(* IEC 61131-3 sources: volt/packages/volt-lsp-iec/test-corpus/bakon-nano/Device/Plc Logic/Application/Library Manager/L_MC1P_MotionControlBasic (part 2) *)

(* ---- L_MC1P_IAXISCOMMMAND.itf ---- *)
INTERFACE L_MC1P_IAXISCOMMMAND
END_INTERFACE

METHOD ABORTING
END_METHOD

METHOD CALCSTATUS
VAR_IN_OUT
	AXIS : _AXIS_REF_REAL;
END_VAR
END_METHOD

METHOD EXECUTE
END_METHOD

METHOD MAIN
END_METHOD

METHOD RESETCOMMANDERRORSTATE : BOOL
VAR_IN_OUT
	AXIS : _AXIS_REF_REAL;
END_VAR
END_METHOD

METHOD RESETSTATUSPARAMETER
END_METHOD

METHOD SETINCTANCEINFO
VAR_INPUT
	PSINSTANCENAME : POINTER TO STRING;
	ERRORITFID : DWORD;
END_VAR
END_METHOD

METHOD UPDATEAXISPOINTER
VAR_INPUT
	PAXIS : POINTER TO AXIS_REF;
END_VAR
END_METHOD

METHOD UPDATECOMMANDINTERFACE
VAR_IN_OUT
	CMD : USINT;
END_VAR
END_METHOD

(* ---- L_MC1P_IAXISCOMMMAND_AUTOTUNING.itf ---- *)
INTERFACE L_MC1P_IAXISCOMMMAND_AUTOTUNING
END_INTERFACE

METHOD CALCPROFILEPARAMS
VAR_IN_OUT
	AXIS : AXIS_REF;
END_VAR
END_METHOD

METHOD UPDATEPARAINTERFACE
VAR_IN_OUT
	SCPAR : L_MC1P_AutotuningPara;
END_VAR
END_METHOD

(* ---- L_MC1P_IAXISEXTENSION.itf ---- *)
INTERFACE L_MC1P_IAXISEXTENSION
END_INTERFACE

METHOD SETBASICINITIALISATION
VAR_INPUT
	ITFGENERICCONFIG : L_MC1P_IGenericAxisConfiguration;
END_VAR
VAR_IN_OUT
	AXIS : _AXIS_REF_REAL;
END_VAR
END_METHOD

(* ---- L_MC1P_IAXISSIMCALLSINGLESTEPS.itf ---- *)
INTERFACE L_MC1P_IAXISSIMCALLSINGLESTEPS
END_INTERFACE

METHOD SIMFINISH : BOOL
VAR_INPUT
	AXISID : INT;
	ITFMECHANICSIMULATION : L_MC1P_IMechanicSimulation;
END_VAR
VAR_IN_OUT
	AXIS : _AXIS_REF_REAL;
END_VAR
END_METHOD

METHOD SIMINSIDELOOP : BOOL
VAR_INPUT
	AXISID : INT;
	ISYSTEMSIMCOUNTER : INT;
	ITFMECHANICSIMULATION : L_MC1P_IMechanicSimulation;
END_VAR
END_METHOD

METHOD SIMPREPARE : BOOL
VAR_INPUT
	AXISID : INT;
	ITFMECHANICSIMULATION : L_MC1P_IMechanicSimulation;
END_VAR
VAR_IN_OUT
	AXIS : _AXIS_REF_REAL;
END_VAR
END_METHOD

(* ---- L_MC1P_IAXISSIMULATIONINTERFACE.itf ---- *)
INTERFACE L_MC1P_IAXISSIMULATIONINTERFACE
END_INTERFACE

METHOD ACTIVATESIMULATION
VAR_IN_OUT
	AXIS : _AXIS_REF_REAL;
END_VAR
END_METHOD

METHOD CALCULATEINPUTDATA
VAR_INPUT
	ITFKINSIM : L_MC1P_IKinematicSimulation;
END_VAR
VAR_IN_OUT
	AXIS : _AXIS_REF_REAL;
END_VAR
END_METHOD

METHOD CALCULATEOUTPUTDATA
VAR_INPUT
	ITFKINSIM : L_MC1P_IKinematicSimulation;
END_VAR
VAR_IN_OUT
	AXIS : _AXIS_REF_REAL;
END_VAR
END_METHOD

METHOD DISABLESIMULATION
VAR_IN_OUT
	AXIS : _AXIS_REF_REAL;
END_VAR
END_METHOD

(* ---- L_MC1P_ICOMMMUNICATIONSIMULATION.itf ---- *)
INTERFACE L_MC1P_ICOMMMUNICATIONSIMULATION
END_INTERFACE

METHOD GETCOMMSTATE : L_DCO_CommState
VAR_INPUT
	PAXISCOMM : POINTER TO _AXIS_REF_COM;
END_VAR
END_METHOD

METHOD PARREAD
VAR_INPUT
	WIDX : DWORD;
END_VAR
END_METHOD

METHOD PARREAD_GETOUTPUT
VAR_INPUT
	WIDX : DWORD;
END_VAR
VAR_OUTPUT
	SZDATAREAD : CAA_SIZE;
	XDONE : BOOL;
	XERROR : BOOL;
	WERROR : WORD;
END_VAR
END_METHOD

METHOD PARREAD_SETINPUT
VAR_INPUT
	WIDX : DWORD;
	XEXECUTE : BOOL;
	WINDEX : WORD;
	BYSUBINDEX : BYTE;
	PBUFFER : POINTER TO BYTE;
	SZSIZE : UDINT;
	UDITIMEOUT : UDINT;
	XSLOTB : BOOL;
END_VAR
END_METHOD

METHOD PARWRITE
VAR_INPUT
	WIDX : DWORD;
END_VAR
END_METHOD

METHOD PARWRITE_GETOUTPUT
VAR_INPUT
	WIDX : DWORD;
END_VAR
VAR_OUTPUT
	XDONE : BOOL;
	XERROR : BOOL;
	WERROR : WORD;
END_VAR
END_METHOD

METHOD PARWRITE_SETINPUT
VAR_INPUT
	WIDX : DWORD;
	XEXECUTE : BOOL;
	WINDEX : WORD;
	BYSUBINDEX : BYTE;
	PBUFFER : POINTER TO BYTE;
	SZSIZE : UDINT;
	UDITIMEOUT : UDINT;
	XSLOTB : BOOL;
END_VAR
END_METHOD

METHOD RESTARTMASTER
VAR_INPUT
	XEXECUTE : BOOL;
	PAXIS : POINTER TO _AXIS_REF_COM;
END_VAR
VAR_OUTPUT
	XDONE : BOOL;
	XERROR : BOOL;
	XBUSY : BOOL;
	DWERROR : DWORD;
END_VAR
END_METHOD

(* ---- L_MC1P_ICOMMUNICATION.itf ---- *)
INTERFACE L_MC1P_ICOMMUNICATION
END_INTERFACE

METHOD FORWARDERROR
VAR_INPUT
	XENABLE : BOOL;
	XWARNING : BOOL;
	XERROR : BOOL;
	WERRORID : WORD;
	WTEXTREFID : WORD;
	XRESETERROR : BOOL := FALSE;
	AXISMODULEHANDLER : L_IMHP_IModuleHandler;
END_VAR
END_METHOD

METHOD GETCOMMPARAMETER
VAR_INPUT
	PCONNECTOR : POINTER TO IoConfigConnector;
END_VAR
VAR_OUTPUT
	PSLAVECONNECTOR : POINTER TO IoStandard.IoConfigConnector;
	UINETID : UINT;
	UIDEVICEID : UINT;
	XSENDFRAMEATTASKSTART : BOOL;
	UDIPRODUCTCODE : DWORD;
	PMASTERCONNECTOR : POINTER TO IoStandard.IoConfigConnector;
END_VAR
END_METHOD

METHOD GETCOMMSTATE : L_DCO_CommState
VAR_INPUT
	PAXISCOMM : POINTER TO _AXIS_REF_COM;
END_VAR
END_METHOD

METHOD GETPDINEQPDOUT : BOOL
END_METHOD

METHOD PARREAD
VAR_INPUT
	WIDX : DWORD;
END_VAR
END_METHOD

METHOD PARREAD_GETOUTPUT
VAR_INPUT
	WIDX : DWORD;
END_VAR
VAR_OUTPUT
	SZDATAREAD : CAA_SIZE;
	XDONE : BOOL;
	XERROR : BOOL;
	WERROR : WORD;
END_VAR
END_METHOD

METHOD PARREAD_SETINPUT
VAR_INPUT
	WIDX : DWORD;
	XEXECUTE : BOOL;
	WINDEX : WORD;
	BYSUBINDEX : BYTE;
	PBUFFER : POINTER TO BYTE;
	SZSIZE : UDINT;
	UDITIMEOUT : UDINT;
END_VAR
END_METHOD

METHOD PARWRITE
VAR_INPUT
	WIDX : DWORD;
END_VAR
END_METHOD

METHOD PARWRITE_GETOUTPUT
VAR_INPUT
	WIDX : DWORD;
END_VAR
VAR_OUTPUT
	XDONE : BOOL;
	XERROR : BOOL;
	WERROR : WORD;
END_VAR
END_METHOD

METHOD PARWRITE_SETINPUT
VAR_INPUT
	WIDX : DWORD;
	XEXECUTE : BOOL;
	WINDEX : WORD;
	BYSUBINDEX : BYTE;
	PBUFFER : POINTER TO BYTE;
	SZSIZE : UDINT;
	UDITIMEOUT : UDINT;
END_VAR
END_METHOD

METHOD RESET
END_METHOD

METHOD RESTARTMASTER
VAR_INPUT
	XEXECUTE : BOOL;
	PAXIS : POINTER TO _AXIS_REF_COM;
END_VAR
VAR_OUTPUT
	XDONE : BOOL;
	XERROR : BOOL;
	XBUSY : BOOL;
	DWERROR : DWORD;
END_VAR
END_METHOD

METHOD SETBASICINITIALISATION
VAR_IN_OUT
	AXIS : _AXIS_REF_REAL;
END_VAR
END_METHOD

METHOD SETCOMPONENTINFO
VAR_INPUT
	DATASELECTION : WORD;
	SDATA : STRING;
END_VAR
END_METHOD

(* ---- L_MC1P_ICOMPENSATIONINTERFACE.itf ---- *)
INTERFACE L_MC1P_ICOMPENSATIONINTERFACE
END_INTERFACE

METHOD GETOFFSETVALUES
VAR_OUTPUT
	LROFFSETPOS : LREAL;
	LROFFSETVEL : LREAL;
	LROFFSETACC : LREAL;
END_VAR
END_METHOD

(* ---- L_MC1P_ICONFIGUREDRIVE.itf ---- *)
INTERFACE L_MC1P_ICONFIGUREDRIVE
END_INTERFACE

METHOD DOFUNCTION : BOOL
VAR_INPUT
	XEXECUTE : BOOL;
	WOFFSET : WORD;
END_VAR
VAR_OUTPUT
	XDONE : BOOL;
	XERROR : BOOL;
	XBUSY : BOOL;
	EERRORID : WORD;
END_VAR
VAR_IN_OUT
	AXIS : _AXIS_REF_REAL;
END_VAR
END_METHOD

METHOD GETADDITIONALCONFIGINFO : POINTER TO L_MC1P_AdditionalConfigInfo
END_METHOD

METHOD GETINSTANCE : POINTER TO BYTE
END_METHOD

METHOD RESET : BOOL
END_METHOD

(* ---- L_MC1P_ICONTROLLERADAPTION.itf ---- *)
INTERFACE L_MC1P_ICONTROLLERADAPTION
END_INTERFACE

METHOD CALCADAPTIONCURVE : LREAL
VAR_INPUT
	LRSETVEL : LREAL;
END_VAR
VAR_IN_OUT
	AXIS : _AXIS_REF_REAL;
END_VAR
END_METHOD

(* ---- L_MC1P_ICONTROLLERINTERFACE.itf ---- *)
INTERFACE L_MC1P_ICONTROLLERINTERFACE
END_INTERFACE

METHOD CALCCONTROLLER
VAR_INPUT
	LRSETPOSITION : LREAL;
	LRSETVELOCITY : LREAL;
	LRSETACCELERATION : LREAL;
	LRSETTORQUE : LREAL;
	LRSETJERK : LREAL;
	LRACTPOSITIONIN : LREAL;
	LRACTVELOCITYIN : LREAL;
	LRACTACCELERATIONIN : LREAL;
	LRACTTORQUEIN : LREAL;
END_VAR
VAR_OUTPUT
	LRSETPOSITIONOUT : LREAL;
	LRSETVELOCITYOUT : LREAL;
	LRSETACCELERATIONOUT : LREAL;
	LRSETTORQUEOUT : LREAL;
END_VAR
VAR_IN_OUT
	AXIS : _AXIS_REF_REAL;
END_VAR
END_METHOD

(* ---- L_MC1P_IDRIVESCALING.itf ---- *)
INTERFACE L_MC1P_IDRIVESCALING
END_INTERFACE

METHOD CALCACCFACTOR : BOOL
VAR_OUTPUT
	LRSCALEUNITTOACC : LREAL;
	LRSCALEACCTOUNIT : LREAL;
END_VAR
VAR_IN_OUT
	AXIS : _AXIS_REF_REAL;
END_VAR
END_METHOD

METHOD CALCSPEEDFACTOR : BOOL
VAR_OUTPUT
	LRSCALEUNITTOSPEED : LREAL;
	LRSCALESPEEDTOUNIT : LREAL;
END_VAR
VAR_IN_OUT
	AXIS : _AXIS_REF_REAL;
END_VAR
END_METHOD

METHOD CALCTORQUEFACTOR : BOOL
VAR_OUTPUT
	LRSCALETORQUETONORM : LREAL;
	LRSCALETORQUETONORM2 : LREAL;
	LRSCALENORMTOTORQUE : LREAL;
END_VAR
VAR_IN_OUT
	AXIS : _AXIS_REF_REAL;
END_VAR
END_METHOD

METHOD CHECKVALIDPOSRESOLUTION : BOOL
VAR_INPUT
	DWPOSRESOLUTION : DWORD;
END_VAR
END_METHOD

METHOD GETDEFAULTTORQUE : LREAL
VAR_INPUT
	LRREFTORQUE : LREAL;
END_VAR
END_METHOD

METHOD POSDIFFTOSPEEDINC : DINT
VAR_INPUT
	DIPOSDIFF : DINT := 0;
	DWFACTOR : DWORD := 1000;
END_VAR
VAR_IN_OUT
	AXIS : _AXIS_REF_REAL;
END_VAR
END_METHOD

METHOD SPEEDTOPOSDIFFINC : DINT
VAR_INPUT
	DISPEED : DINT := 0;
	DWFACTOR : DWORD := 1000;
END_VAR
VAR_IN_OUT
	AXIS : _AXIS_REF_REAL;
	DIRES : DINT;
END_VAR
END_METHOD

(* ---- L_MC1P_IDRIVESPECIFICIMPLBASE.itf ---- *)
INTERFACE L_MC1P_IDRIVESPECIFICIMPLBASE
END_INTERFACE

METHOD CALCAFTERREADINPUTS
VAR_IN_OUT
	AXIS : _AXIS_REF_REAL;
END_VAR
END_METHOD

METHOD CALCBEFOREREADINPUTS
VAR_IN_OUT
	AXIS : _AXIS_REF_REAL;
END_VAR
END_METHOD

METHOD CALCBEFOREWRITEOUTPUTS
VAR_IN_OUT
	AXIS : _AXIS_REF_REAL;
END_VAR
END_METHOD

METHOD CHECKAVAILABLECONTROLMODE : BOOL
VAR_IN_OUT
	AXIS : _AXIS_REF_REAL;
	POSCTRLDRIVEAVAILABLE : L_IE1P_Error;
	POSCTRLPLCAVAILABLE : L_IE1P_Error;
	SPEEDCTRLDRIVEAVAILABLE : L_IE1P_Error;
	TORQUECTRLDRIVE : L_IE1P_Error;
END_VAR
END_METHOD

METHOD CHECKRESETHOMEPOS
VAR_INPUT
	WFDBSTATUSWORD : WORD;
END_VAR
VAR_IN_OUT
	AXIS : _AXIS_REF_REAL;
END_VAR
END_METHOD

METHOD CHECKSAFETYOPTIONAVAILABLE : BOOL
VAR_INPUT
	DWPRODUCTCODE : DWORD;
END_VAR
END_METHOD

METHOD COLLECTDRIVESTATE : BOOL
VAR_IN_OUT
	AXIS : _AXIS_REF_REAL;
	SCSTATEINFO : L_MC1P_DriveStateCollection;
END_VAR
END_METHOD

METHOD CONTROLDRIVE : BOOL
VAR_INPUT
	XENABLE : BOOL;
END_VAR
VAR_IN_OUT
	AXIS : _AXIS_REF_REAL;
END_VAR
END_METHOD

METHOD DRIVECONFIGDATA
VAR_INPUT
	PCONFIGINFO : POINTER TO L_MC1P_AdditionalConfigInfo;
END_VAR
VAR_IN_OUT
	AXIS : _AXIS_REF_REAL;
END_VAR
END_METHOD

METHOD DRIVEFAULTSTATUS : BOOL
VAR_IN_OUT
	AXIS : _AXIS_REF_REAL;
	SCSTATEINFO : L_MC1P_DriveStateCollection;
END_VAR
END_METHOD

METHOD GETBRAKE : POINTER TO L_MC1P_BrakeControlBase
VAR_IN_OUT
	AXIS : _AXIS_REF_REAL;
END_VAR
END_METHOD

METHOD GETBRAKESERVICE : POINTER TO L_MC1P_BrakeService
VAR_IN_OUT
	AXIS : _AXIS_REF_REAL;
END_VAR
END_METHOD

METHOD GETCAUSEOFCINH : WORD
VAR_IN_OUT
	AXIS : _AXIS_REF_REAL;
END_VAR
END_METHOD

METHOD GETFDBSTATUSWORD : WORD
VAR_IN_OUT
	AXIS : _AXIS_REF_REAL;
END_VAR
END_METHOD

METHOD GETIECADRESS : BOOL
VAR_IN_OUT
	AXIS : _AXIS_REF_REAL;
	M_PPDOINFOCONNECTOR : POINTER TO IoConfigConnector;
	ATRANSELEMENT : ARRAY [1.._AXIS_REF_REAL.c_wMaxTransElem] OF L_MC1P_MappedElement;
	WTRANSELEMENTS : WORD;
	LWTRANSDATA : LWORD;
	LWRECDATA : LWORD;
	WRECEIVEELEMENTS : WORD;
	ARECEIVEELEMENT : ARRAY [1.._AXIS_REF_REAL.c_wMaxRecElem] OF L_MC1P_MappedElement;
END_VAR
END_METHOD

METHOD GETOPTIONALACTVEL : BOOL
VAR_IN_OUT
	LRVEL : LREAL;
END_VAR
END_METHOD

METHOD GETRECEIVEDATAIMPL : DWORD
VAR_INPUT
	LWMASK : LWORD;
END_VAR
VAR_IN_OUT
	AXIS : _AXIS_REF_REAL;
END_VAR
END_METHOD

METHOD GETSTATUSWORDS
VAR_OUTPUT
	STATUSWORD1 : WORD;
	STATUSWORD2 : WORD;
	STATUSWORD3 : WORD;
	STATUSWORD4 : WORD;
END_VAR
VAR_IN_OUT
	AXIS : _AXIS_REF_REAL;
END_VAR
END_METHOD

METHOD GETTRANSMITDATAIMPL : DWORD
VAR_INPUT
	LWMASK : LWORD;
END_VAR
VAR_IN_OUT
	AXIS : _AXIS_REF_REAL;
END_VAR
END_METHOD

METHOD GETTRANSMITDATALREALIMPL : LREAL
VAR_INPUT
	LWMASK : LWORD;
END_VAR
VAR_IN_OUT
	AXIS : _AXIS_REF_REAL;
END_VAR
END_METHOD

METHOD HOMECONFIG : BOOL
VAR_INPUT
	LRPOSITION : LREAL;
END_VAR
VAR_OUTPUT
	WINDEX : WORD;
	BYSUBINDEX : BYTE;
	BYNROFBYTE : BYTE;
	DWDATA : DWORD;
	XWRITEPARAM : BOOL;
	XDONE : BOOL;
	XERROR : BOOL;
END_VAR
VAR_IN_OUT
	AXIS : _AXIS_REF_REAL;
	SCHOMEDATA : L_MC1P_HomeParameter;
	WSTEP : WORD;
END_VAR
END_METHOD

METHOD HOMEPOSPERMANENTSETACTIVE : BOOL
VAR_IN_OUT
	AXIS : _AXIS_REF_REAL;
END_VAR
END_METHOD

METHOD RECEIVEPARAMETER
VAR_INPUT
	WPARAMETER : WORD;
	PADRESS : POINTER TO BYTE;
	WSIZE : WORD;
END_VAR
VAR_IN_OUT
	AXIS : _AXIS_REF_REAL;
END_VAR
END_METHOD

METHOD RECEIVEPARAMETERCALC
VAR_IN_OUT
	AXIS : _AXIS_REF_REAL;
	DATA : ARRAY [1..L_MC1P_Constants.gc_Rec_MaxDataIndex] OF POINTER TO L_MC1P_MappedElement;
END_VAR
END_METHOD

METHOD RESETDRIVECONTROL
VAR_INPUT
	XRESETDRIVEERROR : BOOL;
END_VAR
END_METHOD

METHOD RESTOREADDITIONALRETAINDATA
VAR_INPUT
	PDATA : POINTER TO L_MC1P_uRetainData;
END_VAR
END_METHOD

METHOD SETAXISPROPERTIES
VAR_IN_OUT
	AXIS : _AXIS_REF_REAL;
	AXISPROPERTIES : L_MC1P_AxisProperties;
END_VAR
END_METHOD

METHOD SETAXISSTATUSWORD
VAR_IN_OUT
	AXIS : _AXIS_REF_REAL;
	DWAXISSTATUS : DWORD;
END_VAR
END_METHOD

METHOD SETBASICINITIALISATION
VAR_IN_OUT
	AXIS : _AXIS_REF_REAL;
END_VAR
END_METHOD

METHOD SETCONTROLWORDS
VAR_INPUT
	CONTROLWORD1 : WORD;
	CONTROLWORD2 : WORD;
	CONTROLWORD3 : WORD;
	CONTROLWORD4 : WORD;
END_VAR
VAR_IN_OUT
	AXIS : _AXIS_REF_REAL;
END_VAR
END_METHOD

METHOD SETDCBRAKE
VAR_INPUT
	XSETDCBRAKE : BOOL;
END_VAR
VAR_OUTPUT
	XDCBRAKEACTIVE : BOOL;
END_VAR
VAR_IN_OUT
	AXIS : _AXIS_REF_REAL;
END_VAR
END_METHOD

METHOD SETDRIVECONFIGINIT
VAR_IN_OUT
	AXIS : _AXIS_REF_REAL;
END_VAR
END_METHOD

METHOD SETSPEEDCTRLLIMITATION : BOOL
VAR_INPUT
	XLIMIT : BOOL;
END_VAR
VAR_IN_OUT
	AXIS : _AXIS_REF_REAL;
END_VAR
END_METHOD

METHOD SETSPEEDCTRLLOADVALUE
VAR_INPUT
	XLOAD : BOOL;
	LRVALUE : LREAL;
END_VAR
VAR_IN_OUT
	AXIS : _AXIS_REF_REAL;
END_VAR
END_METHOD

METHOD STOREADDITIONALRETAINDATA
VAR_INPUT
	PDATA : POINTER TO L_MC1P_uRetainData;
END_VAR
END_METHOD

METHOD TRANSMITPARAMETER
VAR_INPUT
	WPARAMETER : WORD;
	PADRESS : POINTER TO BYTE;
	WSIZE : WORD;
END_VAR
VAR_IN_OUT
	AXIS : _AXIS_REF_REAL;
END_VAR
END_METHOD

METHOD TRANSMITPARAMETERCALC
VAR_IN_OUT
	AXIS : _AXIS_REF_REAL;
	DATA : ARRAY [1..L_MC1P_Constants.gc_Trans_MaxDataIndex] OF POINTER TO L_MC1P_MappedElement;
END_VAR
END_METHOD

METHOD UPDATEMAPPING
VAR_INPUT
	PTASKMAPLIST : POINTER TO IoStandard.IoConfigTaskMap;
	NCOUNT : DINT;
	PPDOINFOCONNECTOR : POINTER TO IoConfigConnector;
END_VAR
VAR_IN_OUT
	AXIS : _AXIS_REF_REAL;
END_VAR
END_METHOD

(* ---- L_MC1P_IDRIVEUTILS.itf ---- *)
INTERFACE L_MC1P_IDRIVEUTILS
END_INTERFACE

METHOD ACTIVATEAPPCREDITS
VAR_INPUT
	XACTIVATE : BOOL;
END_VAR
END_METHOD

METHOD GETMULTIAXISINFO
VAR_IN_OUT
	MULTIAXISINFO : L_MC1P_MultiAxisInfo;
END_VAR
END_METHOD

METHOD GETRETAINMEMINFO : L_MC1P_RetainDataType
VAR_OUTPUT
	MEMINFO : L_MC1P_uAxisRetainInfo;
END_VAR
END_METHOD

METHOD RESETCONNECTION : L_IE1P_Error
VAR_INPUT
	ITFCALLEDFUNCITON : L_IF1P_IFunctionConnection;
	EDISCONNECTMODE : L_IF1P_DisconnectMode;
	XDISCONNECTEXISTINGCONNECTION : BOOL;
END_VAR
END_METHOD

METHOD SETCONNECTION
VAR_INPUT
	AXISCONNECTION : L_IF1P_IFunctionConnection;
END_VAR
END_METHOD

(* ---- L_MC1P_IENCODERINTERFACE.itf ---- *)
INTERFACE L_MC1P_IENCODERINTERFACE
END_INTERFACE

METHOD ENCNEWHOMEPOSLOADED : BOOL
VAR_INPUT
	DWCALLYCLE : DWORD;
	DWDELAY : DWORD;
END_VAR
END_METHOD

METHOD ENCRESETACTPOS
END_METHOD

METHOD ENCRESETHOMEPOS
VAR_INPUT
	ERESETINFO : L_IE1P_Error;
END_VAR
END_METHOD

METHOD ENCSETHOMEPOSITION
VAR_INPUT
	POSITION : LREAL;
	RELATIVE : BOOL;
	POSDIFF : LREAL;
	EHOMEPOSINFO : L_IE1P_Error;
END_VAR
END_METHOD

METHOD ENCSIGNALVALID : BOOL
VAR_OUTPUT
	XSIGNALVALIDOLD : BOOL;
	EENCERRORID : L_IE1P_Error;
END_VAR
END_METHOD

METHOD GETACTPOSINCR : DINT
END_METHOD

METHOD GETACTPOSINCR1616 : DINT
END_METHOD

METHOD GETACTVALUES
VAR_OUTPUT
	LRACTPOS : LREAL;
	LRACTVEL : LREAL;
	LRACTACC : LREAL;
	LRACTPOSUNFILTERED : LREAL;
	LRACTPOSROUNDS : LREAL;
END_VAR
END_METHOD

METHOD GETAXISINSTANCE : POINTER TO _AXIS_REF_REAL
END_METHOD

METHOD GETCONFIGCHANGED : BOOL
END_METHOD

METHOD GETHOMEPOSAVAILABLE : BOOL
END_METHOD

METHOD SETHOMEPOSAVAILABLE
VAR_INPUT
	XHOMEPOSAVAILABLE : BOOL;
END_VAR
END_METHOD

(* ---- L_MC1P_IENCODERPOSFILTER.itf ---- *)
INTERFACE L_MC1P_IENCODERPOSFILTER
END_INTERFACE

METHOD CALCULATE
VAR_INPUT
	LRCYCPOSIN : LREAL;
	LRCYCVELIN : LREAL;
END_VAR
VAR_OUTPUT
	LRCYCPOSOUT : LREAL;
	LRCYCVELOUT : LREAL;
	WFILTERSTATE : WORD;
END_VAR
END_METHOD

METHOD INIT
END_METHOD

METHOD RESET
END_METHOD

(* ---- L_MC1P_IERRORHANDLINGAXISSYSTEMS.itf ---- *)
INTERFACE L_MC1P_IERRORHANDLINGAXISSYSTEMS
END_INTERFACE

METHOD CLEARERRORINAXISSYSTEM
VAR_INPUT
	INSTANCEID : DWORD := 0;
END_VAR
END_METHOD

METHOD GETERRORITFID : DWORD
END_METHOD

METHOD NOTIFYERRORINAXISSYSTEM : BOOL
VAR_INPUT
	WERRORID : L_IE1P_Error := 0;
	INSTANCEID : DWORD := 0;
	PSINSTANCENAME : POINTER TO BYTE := 0;
	EERRORREACTION : L_IE1P_SeverityLevel := 0;
END_VAR
END_METHOD

(* ---- L_MC1P_IEXTENDEDMAPPINGACCESS.itf ---- *)
INTERFACE L_MC1P_IEXTENDEDMAPPINGACCESS
END_INTERFACE

METHOD GETIECADRESS
VAR_INPUT
	AXISCONNECTOR : POINTER TO IoConfigConnector;
END_VAR
END_METHOD

METHOD GETMAPPEDDATA : POINTER TO BYTE
VAR_INPUT
	UIINDEX : WORD;
	USISUBINDEX : USINT;
	USISIZE : USINT;
	XWRITEACCESS : BOOL;
	PADDDATA : POINTER TO BYTE;
	PXWAITFORINITACCESS : POINTER TO BOOL;
END_VAR
VAR_OUTPUT
	EERRORID : L_IE1P_Error;
	XERROR : BOOL;
	USISIZEACT : USINT;
END_VAR
END_METHOD

METHOD GETMAPPEDDATASUPPORT : BOOL
END_METHOD

METHOD RESETOUTPUTMAPPINGOBJECTS : BOOL
END_METHOD

(* ---- L_MC1P_IGENERICAXISCONFIGURATION.itf ---- *)
INTERFACE L_MC1P_IGENERICAXISCONFIGURATION
END_INTERFACE

METHOD CALCAFTERREADINPUTS
VAR_IN_OUT
	AXIS : _AXIS_REF_REAL;
	DRIVESPECIFIC : L_MC1P_DriveSpecific_Generic;
END_VAR
END_METHOD

METHOD CALCBEFOREREADINPUTS
VAR_IN_OUT
	AXIS : _AXIS_REF_REAL;
	DRIVESPECIFIC : L_MC1P_DriveSpecific_Generic;
END_VAR
END_METHOD

METHOD CALCBEFOREWRITEOUTPUTS
VAR_IN_OUT
	AXIS : _AXIS_REF_REAL;
	DRIVESPECIFIC : L_MC1P_DriveSpecific_Generic;
END_VAR
END_METHOD

METHOD DRIVECONFIG
VAR_INPUT
	WOFFSET : WORD;
END_VAR
VAR_OUTPUT
	XCONFIGBUSY : BOOL;
	XWAITFORPARAMETERWRITEDONE : BOOL;
	XWAITFORPARAMETERREADDONE : BOOL;
	XREADSTRING : BOOL;
	DWWRITEDATA : DWORD;
	WINDEX : WORD;
	BYSUBINDEX : BYTE;
	BYNROFBYTE : BYTE;
END_VAR
VAR_IN_OUT
	AXIS : _AXIS_REF_REAL;
	CONFIGINFO : L_MC1P_AdditionalConfigInfo;
	WSTEP : WORD;
	EERRORID : WORD;
	DWREADDATA : DWORD;
	SREADDATA : STRING(255);
END_VAR
END_METHOD

METHOD GETADDITIONALSTATEINFOS : BOOL
VAR_IN_OUT
	AXIS : _AXIS_REF_REAL;
	DRIVESPECIFIC : L_MC1P_DriveSpecific_Generic;
	SCSTATEINFO : L_MC1P_DriveStateCollection;
END_VAR
END_METHOD

METHOD GETHOMINGSTATE
VAR_INPUT
	WHOMESTATE : WORD;
END_VAR
VAR_IN_OUT
	AXIS : _AXIS_REF_REAL;
	XHOMEPOSAVAILABLEDRIVE : BOOL;
END_VAR
END_METHOD

METHOD HOMECONFIG
VAR_INPUT
	LRPOSITION : LREAL;
END_VAR
VAR_OUTPUT
	XCONFIGBUSY : BOOL;
	XERROR : BOOL;
	WINDEX : WORD;
	BYSUBINDEX : BYTE;
	BYNROFBYTE : BYTE;
	DWDATA : DWORD;
	XWRITEPARAM : BOOL;
END_VAR
VAR_IN_OUT
	AXIS : _AXIS_REF_REAL;
	SCHOMEDATA : L_MC1P_HomeParameter;
	WSTEP : WORD;
END_VAR
END_METHOD

METHOD RECEIVEPARAMETERCALC
VAR_IN_OUT
	AXIS : _AXIS_REF_REAL;
	DATA : ARRAY [1..L_MC1P_Constants.gc_Rec_MaxDataIndex] OF POINTER TO L_MC1P_MappedElement;
	DRIVESPECIFIC : L_MC1P_DriveSpecific_Generic;
END_VAR
END_METHOD

METHOD TRANSMITPARAMETERCALC
VAR_IN_OUT
	AXIS : _AXIS_REF_REAL;
	DATA : ARRAY [1..L_MC1P_Constants.gc_Trans_MaxDataIndex] OF POINTER TO L_MC1P_MappedElement;
	DRIVESPECIFIC : L_MC1P_DriveSpecific_Generic;
END_VAR
END_METHOD

(* ---- L_MC1P_IKINEMATICMASTER.itf ---- *)
INTERFACE L_MC1P_IKINEMATICMASTER
END_INTERFACE

METHOD ACTIVATEHOMESIGNALMONITORINGSLAVE
END_METHOD

METHOD ADDOFFSETVALUESFORMASTER
VAR_IN_OUT
	LRSETPOSITION : LREAL;
	LRSETVELOCITY : LREAL;
	LRSETACCELERATION : LREAL;
	LRSETTORQUE : LREAL;
END_VAR
END_METHOD

METHOD FINISHHOMINGFORMASTERAXIS : BOOL
END_METHOD

METHOD GETERRORACTIVEMAINAXIS : BOOL
END_METHOD

METHOD GETERRORSETVALUESFROMMAINAXIS : BOOL
VAR_INPUT
	XCONTROLLEDSTOPPOSSIBLE : BOOL;
END_VAR
VAR_OUTPUT
	XSETQSP : BOOL;
	XSETCINH : BOOL;
END_VAR
END_METHOD

METHOD GETMASTERAXISINSTANCE : POINTER TO AXIS_REF
END_METHOD

METHOD SETERRORMAINAXIS : BOOL
VAR_INPUT
	ESEVERITY : L_IE1P_SeverityLevel;
	WERRORID : WORD;
	DWEXTENDEDERRORINFO : DWORD;
END_VAR
END_METHOD

METHOD SWITCHROLE : BOOL
VAR_INPUT
	XSWITCH : BOOL;
END_VAR
END_METHOD

METHOD WAITHOMINGFORMASTERAXIS : BOOL
END_METHOD

METHOD FINISHBRAKETESTFORMASTERAXIS : BOOL
END_METHOD

METHOD FINISHGRINDINFORMASTERAXIS : BOOL
END_METHOD

METHOD WAITBRAKETESTFORMASTERAXIS : BOOL
END_METHOD

METHOD WAITGRINDINFORMASTERAXIS : BOOL
END_METHOD

(* ---- L_MC1P_IKINEMATICSIMULATION.itf ---- *)
INTERFACE L_MC1P_IKINEMATICSIMULATION
END_INTERFACE

METHOD CALLSYSSIM : BOOL
VAR_IN_OUT
	AXIS : _AXIS_REF_REAL;
END_VAR
END_METHOD

METHOD INITNEWCYCLE : BOOL
VAR_IN_OUT
	AXIS : _AXIS_REF_REAL;
END_VAR
END_METHOD

METHOD SETAXIS
VAR_INPUT
	AXISID : INT;
	PAXIS : POINTER TO _AXIS_REF_REAL;
END_VAR
END_METHOD

METHOD SETREQUIREDNUMBEROFAXIS
VAR_INPUT
	INUMAXIS : INT;
END_VAR
END_METHOD

(* ---- L_MC1P_IKINEMATICSLAVE.itf ---- *)
INTERFACE L_MC1P_IKINEMATICSLAVE
END_INTERFACE

METHOD ABORTHOMINGSLAVE : BOOL
END_METHOD

METHOD ACTIVATEHOMESIGNALMONITORINGMASTER
END_METHOD

METHOD ACTIVEMASTERHOMEPARAMETER
VAR_INPUT
	EHOMEMODE : L_MC1P_HomeMode;
	LRHOMEPOSITION : LREAL;
END_VAR
END_METHOD

METHOD ADDOFFSETVALUESFORSLAVE
VAR_IN_OUT
	LRSETPOSITION : LREAL;
	LRSETVELOCITY : LREAL;
	LRSETACCELERATION : LREAL;
	LRSETTORQUE : LREAL;
END_VAR
END_METHOD

METHOD CHECKHOMEPARAMETER : BOOL
VAR_OUTPUT
	XERROR : BOOL;
	EERRORID : L_IE1P_Error;
END_VAR
VAR_IN_OUT
	SCHOMEPARAMETER : L_MC1P_HomeParameter;
END_VAR
END_METHOD

METHOD DOHOMINGSLAVE : BOOL
END_METHOD

METHOD FINISHHOMINGFORSLAVEAXIS : BOOL
END_METHOD

METHOD GETERRORACTIVEFOLLOWAXIS : BOOL
END_METHOD

METHOD GETERRORSETVALUESFROMFOLLOWAXIS : BOOL
VAR_INPUT
	XCONTROLLEDSTOPPOSSIBLE : BOOL;
END_VAR
VAR_OUTPUT
	XSETQSP : BOOL;
	XSETCINH : BOOL;
END_VAR
END_METHOD

METHOD GETEXTERNALAUTOTUNINGITF : POINTER TO BYTE
VAR_INPUT
	XRESET : BOOL;
	UIACTUALATNBR : UINT;
END_VAR
VAR_OUTPUT
	WNBOFAUTOTUNINGS : WORD;
END_VAR
END_METHOD

METHOD GETMAXVEL : LREAL
VAR_IN_OUT
	LRVEL : LREAL;
END_VAR
END_METHOD

METHOD GETSETVALUESAVAILABLEMASTER : BOOL
END_METHOD

METHOD GETSLAVEAXISENABLED : BOOL
END_METHOD

METHOD GETSLAVEAXISHOMINGDONE : BOOL
END_METHOD

METHOD GETSLAVEAXISINSTANCE : POINTER TO AXIS_REF
END_METHOD

METHOD MOTIONALLOWED : BOOL
VAR_INPUT
	ETYPEFUNCTION : L_MC1P_TypeFunction;
END_VAR
VAR_OUTPUT
	EERRORCAUSE : L_IE1P_Error;
END_VAR
END_METHOD

METHOD RESETHOMEPOS
VAR_INPUT
	ERESETINFO : L_IE1P_Error;
	XRESETPOSITION : BOOL;
END_VAR
END_METHOD

METHOD RESTOREFOLLOWINGAXISERROR : BOOL
VAR_INPUT
	ESEVERITY : L_IE1P_SeverityLevel;
	WERRORID : WORD;
	DWEXTENDEDERRORINFO : DWORD;
END_VAR
END_METHOD

METHOD SETERRORFOLLOWAXIS : BOOL
VAR_INPUT
	ESEVERITY : L_IE1P_SeverityLevel;
	WERRORID : WORD;
	DWEXTENDEDERRORINFO : DWORD;
END_VAR
END_METHOD

METHOD SETHOMEPOS
VAR_INPUT
	POSITION : LREAL;
	RELATIVE : BOOL;
	XRESTARTPOSITIONING : BOOL := FALSE;
	EHOMEPOSINFO : L_IE1P_Error;
END_VAR
END_METHOD

METHOD SLAVEAXISRESETERROR : BOOL
END_METHOD

METHOD SLAVEAXISRESETPOSSIBLE : BOOL
END_METHOD

METHOD SWITCHROLE : BOOL
VAR_INPUT
	XSWITCH : BOOL;
END_VAR
END_METHOD

METHOD UPDATEABCSTATE : POINTER TO L_MC1P_AxisBasicControlOutput_Internal
END_METHOD

METHOD WAITHOMINGFORSLAVEAXIS : BOOL
END_METHOD

METHOD ABORTBRAKETESTSLAVE : BOOL
VAR_INPUT
	XMAINABORTED : BOOL;
END_VAR
END_METHOD

METHOD DOBRAKETESTSLAVE : BOOL
END_METHOD

METHOD FINISHBRAKETESTFORSLAVEAXIS : BOOL
END_METHOD

METHOD GETBTSTATUS : LREAL
END_METHOD

METHOD GETSLAVEAXISBRAKETESTDONE : BOOL
END_METHOD

METHOD WAITBRAKETESTFORSLAVEAXIS : BOOL
END_METHOD

METHOD ABORTGRINDINSLAVE : BOOL
VAR_INPUT
	XMAINABORTED : BOOL;
END_VAR
END_METHOD

METHOD DOGRINDINSLAVE : BOOL
END_METHOD

METHOD FINISHGRINDINFORSLAVEAXIS : BOOL
END_METHOD

METHOD GETACTIVEGRINDINCYCLESDONE : WORD
VAR_INPUT
	WCYCLESDONE : WORD;
END_VAR
END_METHOD

METHOD GETGICYCLES : LREAL
END_METHOD

METHOD GETGISTATUS : LREAL
END_METHOD

METHOD GETSLAVEAXISGRINDINDONE : BOOL
END_METHOD

METHOD WAITGRINDINFORSLAVEAXIS : BOOL
END_METHOD

(* ---- L_MC1P_ILMDATA.itf ---- *)
INTERFACE L_MC1P_ILMDATA
END_INTERFACE

METHOD ABORT : UDINT
END_METHOD

METHOD EXECUTE : UDINT
END_METHOD

(* ---- L_MC1P_IMANAGEMENTFUNCTION.itf ---- *)
INTERFACE L_MC1P_IMANAGEMENTFUNCTION
END_INTERFACE

METHOD COMPAREAXISNAME : BOOL
VAR_IN_OUT
	SAXISNAME : STRING;
END_VAR
END_METHOD

METHOD GETAXIS : POINTER TO AXIS_REF
END_METHOD

(* ---- L_MC1P_IMANIPULATEACTVALUES.itf ---- *)
INTERFACE L_MC1P_IMANIPULATEACTVALUES
END_INTERFACE

METHOD MANIPULATEACTVALUES
VAR_IN_OUT
	AXIS : AXIS_REF;
END_VAR
END_METHOD

(* ---- L_MC1P_IMANIPULATIONINTERFACE.itf ---- *)
INTERFACE L_MC1P_IMANIPULATIONINTERFACE
END_INTERFACE

METHOD CALCVALUES
VAR_INPUT
	XENABLE : BOOL;
	XRESET : BOOL;
	LRSETPOS : LREAL;
	LRSETVEL : LREAL;
	LRSETACC : LREAL;
	LRSETTORQUE : LREAL;
	XLOADPOSOFFSET : BOOL;
	LRPOSOFFSET : LREAL;
END_VAR
VAR_OUTPUT
	XACTIVE : BOOL;
	XERROR : BOOL;
	EERRORID : L_IE1P.L_IE1P_Error;
	LRSETPOSOUT : LREAL;
	LRSETVELOUT : LREAL;
	LRSETACCOUT : LREAL;
	LRSETTORQUEOUT : LREAL;
END_VAR
VAR_IN_OUT
	AXIS : Axis_REf;
END_VAR
END_METHOD

(* ---- L_MC1P_IMASTERINITINFO.itf ---- *)
INTERFACE L_MC1P_IMASTERINITINFO
END_INTERFACE

(* ---- L_MC1P_IMCPARAMETERACCESS.itf ---- *)
INTERFACE L_MC1P_IMCPARAMETERACCESS
END_INTERFACE

METHOD GETINSTANCEANDTYPE : BOOL
VAR_OUTPUT
	PINSTANCEPOINTER : POINTER TO BYTE;
	EAXISTYPE : L_MC1P_AxisType;
END_VAR
END_METHOD

METHOD HLP_GETPARAMETERPROPERTIES : BOOL
VAR_INPUT
	DIPARAMETER : DINT;
END_VAR
VAR_OUTPUT
	PPARAMADDR : POINTER TO BYTE;
	EORDINALTYPE : L_MC1P_OrdinalType;
	XREADWRITE : BOOL;
	LRUNITFACTOR : LREAL;
	LRDEFAULTVALUE : LREAL;
	WVALUERANGES : WORD;
	PVALUERANGES : POINTER TO L_MC1P_MinMaxValue;
END_VAR
END_METHOD

METHOD HLP_READBOOLPARAMETER : BOOL
VAR_INPUT
	PARAMETER : DINT;
	PXVALUE : POINTER TO BOOL;
END_VAR
END_METHOD

METHOD HLP_READPARAMETER : BOOL
VAR_INPUT
	PARAMETER : DINT;
	PLRVALUE : POINTER TO LREAL;
END_VAR
END_METHOD

METHOD HLP_WRITEBOOLPARAMETER : BOOL
VAR_INPUT
	PARAMETER : DINT;
	PXVALUE : POINTER TO BOOL;
END_VAR
VAR_OUTPUT
	WERRORID : WORD;
END_VAR
END_METHOD

METHOD HLP_WRITEPARAMETER : BOOL
VAR_INPUT
	PARAMETER : DINT;
	PLRVALUE : POINTER TO LREAL;
END_VAR
VAR_OUTPUT
	WERRORID : WORD;
END_VAR
END_METHOD

METHOD QUEUEDPARAMWRITINGACTIVE : BOOL
END_METHOD

(* ---- L_MC1P_IMECHANICSIMULATION.itf ---- *)
INTERFACE L_MC1P_IMECHANICSIMULATION
END_INTERFACE

METHOD CALLMECHANICSIMULATION : BOOL
VAR_INPUT
	AXISID : INT;
	XBRAKERELEASED : BOOL;
	LRACTTORQUE : LREAL;
	LRADDTORQUE : LREAL;
END_VAR
VAR_IN_OUT
	SCPARGENERAL : L_MC1P_ParGeneralMechanic;
END_VAR
END_METHOD

METHOD INITANDSCALEPARAMETER
VAR_INPUT
	AXISID : INT;
	LRTASKCYCLESYSSIM : LREAL;
	LRINVTASKCYCLESYSSIM : LREAL;
END_VAR
VAR_IN_OUT
	SCPARGENERAL : L_MC1P_ParGeneralMechanic;
END_VAR
END_METHOD

METHOD MECHANICSIMGETACTLOADVALUES
VAR_INPUT
	AXISID : INT;
END_VAR
VAR_OUTPUT
	LRACTLOADPOS : LREAL;
	LRACTLOADVEL : LREAL;
END_VAR
END_METHOD

METHOD MECHANICSIMGETACTVALUES
VAR_INPUT
	AXISID : INT;
END_VAR
VAR_OUTPUT
	LRACTPOS : LREAL;
	LRACTVEL : LREAL;
END_VAR
END_METHOD

METHOD SETLOADIDX
VAR_INPUT
	AXISID : INT;
	WIDXLOADMASS : WORD;
END_VAR
END_METHOD

METHOD SETSTARTPOSITION : BOOL
VAR_INPUT
	AXISID : INT;
	LRPOS : LREAL;
END_VAR
END_METHOD

(* ---- L_MC1P_IMOLACCESS.itf ---- *)
INTERFACE L_MC1P_IMOLACCESS
END_INTERFACE

METHOD SETMOLSTATES
VAR_INPUT
	WSETMOLSTATE : WORD := 0;
	WSETMOLMODE : WORD := 0;
END_VAR
END_METHOD

(* ---- L_MC1P_IPARA.itf ---- *)
INTERFACE L_MC1P_IPARA
END_INTERFACE

METHOD HLP_GETPARAMETERPROPERTIES : BOOL
VAR_INPUT
	PAXISREF : POINTER TO AXIS_REF;
	DIPARAMETER : DINT;
	XALLOWINVISIBLE : BOOL;
END_VAR
VAR_OUTPUT
	PPARAMADDR : POINTER TO BYTE;
	EORDINALTYPE : L_MC1P_OrdinalType;
	XREADWRITE : BOOL;
	LRUNITFACTOR : LREAL;
	LRDEFAULTVALUE : LREAL;
	WVALUERANGES : WORD;
	PVALUERANGES : POINTER TO L_MC1P_MinMaxValue;
END_VAR
END_METHOD

METHOD HLP_READBOOLPARAMETER : BOOL
VAR_INPUT
	PINPUTDATA : POINTER TO BYTE;
	PARAMETER : DINT;
	PXVALUE : POINTER TO BOOL;
	XALLOWINVISIBLE : BOOL;
END_VAR
END_METHOD

METHOD HLP_READPARAMETER : BOOL
VAR_INPUT
	PINPUTDATA : POINTER TO BYTE;
	PARAMETER : DINT;
	PLRVALUE : POINTER TO LREAL;
	XALLOWINVISIBLE : BOOL;
END_VAR
END_METHOD

METHOD HLP_WRITEBOOLPARAMETER : BOOL
VAR_INPUT
	PINPUTDATA : POINTER TO BYTE;
	PARAMETER : DINT;
	PXVALUE : POINTER TO BOOL;
	XALLOWINVISIBLE : BOOL;
END_VAR
VAR_OUTPUT
	WERRORID : WORD;
END_VAR
END_METHOD

METHOD HLP_WRITEPARAMETER : BOOL
VAR_INPUT
	PINPUTDATA : POINTER TO BYTE;
	PARAMETER : DINT;
	PLRVALUE : POINTER TO LREAL;
	XALLOWINVISIBLE : BOOL;
END_VAR
VAR_OUTPUT
	WERRORID : WORD;
END_VAR
END_METHOD

(* ---- L_MC1P_IPLIACCESS.itf ---- *)
INTERFACE L_MC1P_IPLIACCESS
END_INTERFACE

METHOD SETPPISTATES
VAR_INPUT
	WSETPPISTATE : WORD := 0;
	WSETPPIMODE : WORD := 0;
END_VAR
END_METHOD

(* ---- L_MC1P_IPOSPROFILECALCULATION.itf ---- *)
INTERFACE L_MC1P_IPOSPROFILECALCULATION
END_INTERFACE

METHOD CALCPROFILEDATA
VAR_INPUT
	PPOSPROFILERDATA : POINTER TO L_MC1P_PosProfiler;
	LRSTARTACC : LREAL;
	LRSTARTVEL : LREAL;
	LRSTARTPOS : LREAL;
	XVELMODE : BOOL;
END_VAR
VAR_OUTPUT
	XERROR : BOOL;
	DWSTATE : DWORD;
	DWPROFILETYPE : DWORD;
END_VAR
VAR_IN_OUT
	SCPROFILEDATA : L_MC1P_ProfileData;
	SCPROFILEPARAMETER : L_MC1P_ProfileParameter;
END_VAR
END_METHOD

METHOD PROFILEINTERPOLATOR : BOOL
VAR_INPUT
	PPOSPROFILERDATA : POINTER TO L_MC1P_PosProfiler;
	LREVALTIME : LREAL;
END_VAR
VAR_OUTPUT
	DWSTATE : DWORD;
	LRSETPOS : LREAL;
	LRSETVEL : LREAL;
	LRSETACC : LREAL;
END_VAR
VAR_IN_OUT
	SCPROFILEDATA : L_MC1P_ProfileData;
END_VAR
END_METHOD

METHOD STRETCHPROFILE
VAR_INPUT
	PPOSPROFILERDATA : POINTER TO L_MC1P_PosProfiler;
	LRTIMEBASE : LREAL;
END_VAR
VAR_IN_OUT
	SCPROFILEDATA : L_MC1P_ProfileData;
END_VAR
END_METHOD

(* ---- L_MC1P_IPOSPROFILERACTIVE.itf ---- *)
INTERFACE L_MC1P_IPOSPROFILERACTIVE
END_INTERFACE

(* ---- L_MC1P_IPOSSIGNALPROCESSING.itf ---- *)
INTERFACE L_MC1P_IPOSSIGNALPROCESSING
END_INTERFACE

METHOD CALCULATE : DINT
VAR_INPUT
	DIACTPOS : DINT;
	DWSAMPLETIME : DWORD;
	DWACTTIME : DWORD;
END_VAR
VAR_OUTPUT
	DIPOSOUT : DINT;
	XVELVALID : BOOL;
	DIVELOUT : DINT;
END_VAR
VAR_IN_OUT
	AXIS : _AXIS_REF_REAL;
END_VAR
END_METHOD

(* ---- L_MC1P_IRETAINFUNCTION.itf ---- *)
INTERFACE L_MC1P_IRETAINFUNCTION
END_INTERFACE

METHOD GETINITIALDATA : BOOL
VAR_INPUT
	PDATA : POINTER TO DWORD;
	INFO : DWORD;
END_VAR
END_METHOD

METHOD SETERRORINFO
VAR_INPUT
	WSTATE : WORD;
END_VAR
END_METHOD

METHOD SETINITIALDATA : BOOL
VAR_INPUT
	PDATA : POINTER TO DWORD;
END_VAR
END_METHOD

METHOD STOREDATA
VAR_INPUT
	PDATA : POINTER TO DWORD;
END_VAR
END_METHOD

(* ---- L_MC1P_IRETAINHANDLING.itf ---- *)
INTERFACE L_MC1P_IRETAINHANDLING
END_INTERFACE

METHOD GETINITIALRETAINDATA : POINTER TO L_MC1P_uRetainData
VAR_INPUT
	XNEWEST : BOOL;
END_VAR
END_METHOD

METHOD GETRETAINSTATE : WORD
VAR_OUTPUT
	WSTATERETAINERROR : WORD;
END_VAR
END_METHOD

METHOD REGISTERONRETAINDATAHANDLER
VAR_INPUT
	AXISGUID : L_MC1P_AxisGUID;
END_VAR
END_METHOD

METHOD RESET
END_METHOD

METHOD SETCONNECTEDGUID : BOOL
VAR_INPUT
	GUID : L_MC1P_AxisGUID;
END_VAR
END_METHOD

(* ---- L_MC1P_ISETSETVALUEMANIPULATORCUSTOM.itf ---- *)
INTERFACE L_MC1P_ISETSETVALUEMANIPULATORCUSTOM
END_INTERFACE

METHOD CALCULATE : L_IE1P_Error
VAR_INPUT
	UIINPUTDATAIDX : UINT;
	UIOUTPUTDATAIDX : UINT;
END_VAR
VAR_IN_OUT
	AXIS : AXIS_REF;
	LRSETPOS : LREAL;
	LRSETVEL : LREAL;
	LRSETACC : LREAL;
	LRSETTORQUE : LREAL;
END_VAR
END_METHOD

METHOD CALLCYCLIC : L_IE1P_Error
VAR_INPUT
	UIINPUTDATAIDX : UINT;
	UIOUTPUTDATAIDX : UINT;
END_VAR
VAR_IN_OUT
	AXIS : Axis_REf;
END_VAR
END_METHOD

METHOD CHECKINPUTDATA : L_IE1P_Error
VAR_INPUT
	UIINPUTDATAIDX : UINT;
	UIOUTPUTDATAIDX : UINT;
END_VAR
VAR_IN_OUT
	AXIS : AXIS_REF;
END_VAR
END_METHOD

METHOD ENABLEEXIT : L_IE1P_Error
VAR_INPUT
	UIINPUTDATAIDX : UINT;
	UIOUTPUTDATAIDX : UINT;
END_VAR
VAR_IN_OUT
	AXIS : AXIS_REF;
END_VAR
END_METHOD

METHOD ENABLEINIT : L_IE1P_Error
VAR_INPUT
	UIINPUTDATAIDX : UINT;
	UIOUTPUTDATAIDX : UINT;
END_VAR
VAR_IN_OUT
	AXIS : AXIS_REF;
END_VAR
END_METHOD

METHOD FREEZEINPUTPERCYCLE
VAR_INPUT
	UIINPUTDATAIDX : UINT;
END_VAR
END_METHOD

METHOD LOADOFFSET : L_IE1P_Error
VAR_INPUT
	UIINPUTDATAIDX : UINT;
	UIOUTPUTDATAIDX : UINT;
	OFFSET : LREAL;
END_VAR
VAR_IN_OUT
	AXIS : Axis_REf;
END_VAR
END_METHOD

METHOD PASSOUTPUTPERCYCLE
VAR_INPUT
	UIOUTPUTDATAIDX : UINT;
END_VAR
END_METHOD

METHOD READINPUTS : L_IE1P_Error
VAR_INPUT
	UIINPUTDATAIDX : UINT;
END_VAR
VAR_IN_OUT
	AXIS : Axis_REf;
END_VAR
END_METHOD

METHOD RESET : L_IE1P_Error
VAR_INPUT
	UIINPUTDATAIDX : UINT;
	UIOUTPUTDATAIDX : UINT;
END_VAR
VAR_IN_OUT
	AXIS : AXIS_REF;
END_VAR
END_METHOD

METHOD RESETOUTPUTS : L_IE1P_Error
VAR_INPUT
	UIOUTPUTDATAIDX : UINT;
END_VAR
VAR_IN_OUT
	AXIS : AXIS_REF;
END_VAR
END_METHOD

(* ---- L_MC1P_ISETVALUEMANIPULATIONINTERFACE.itf ---- *)
INTERFACE L_MC1P_ISETVALUEMANIPULATIONINTERFACE
END_INTERFACE

(* ---- L_MC1P_ITOUCHPROBEHANDLER.itf ---- *)
INTERFACE L_MC1P_ITOUCHPROBEHANDLER
END_INTERFACE

METHOD GETACTTPRECEIVEDATA : L_MC1P_TpReceiveData
END_METHOD

METHOD ISUPTODATE : BOOL
VAR_INPUT
	DWUPDATETIME : DWORD;
END_VAR
END_METHOD

METHOD RECDATAISVALID : BOOL
VAR_IN_OUT
	SCRECDATA : L_MC1P_TpReceiveData;
END_VAR
END_METHOD

(* ---- L_MC1P_ITPSOURCEAXIS.itf ---- *)
INTERFACE L_MC1P_ITPSOURCEAXIS
END_INTERFACE

METHOD GETPOINTERTOTPAXIS : POINTER TO _AXIS_REF_REAL
END_METHOD

(* ---- GETBOOLEANPROPERTY.pou ---- *)
FUNCTION GETBOOLEANPROPERTY : BOOL
VAR_INPUT
	STKEY : WSTRING;
END_VAR
END_FUNCTION

(* ---- GETCOMPANY.pou ---- *)
FUNCTION GETCOMPANY : WSTRING
END_FUNCTION

(* ---- GETNUMBERPROPERTY.pou ---- *)
FUNCTION GETNUMBERPROPERTY : DINT
VAR_INPUT
	STKEY : WSTRING;
END_VAR
END_FUNCTION

(* ---- GETTEXTPROPERTY.pou ---- *)
FUNCTION GETTEXTPROPERTY : WSTRING
VAR_INPUT
	STKEY : WSTRING;
END_VAR
END_FUNCTION

(* ---- GETTEXTPROPERTY2.pou ---- *)
FUNCTION GETTEXTPROPERTY2 : POINTER TO WSTRING
VAR_INPUT
	STKEY : WSTRING;
END_VAR
END_FUNCTION

(* ---- GETTITLE.pou ---- *)
FUNCTION GETTITLE : WSTRING
END_FUNCTION

(* ---- GETVERSION.pou ---- *)
FUNCTION GETVERSION : VERSION
END_FUNCTION

(* ---- GETVERSIONPROPERTY.pou ---- *)
FUNCTION GETVERSIONPROPERTY : VERSION
VAR_INPUT
	STKEY : WSTRING;
END_VAR
END_FUNCTION

(* ---- L_MC1P_CHECKFORSENSORLESMODEIXXX.pou ---- *)
FUNCTION L_MC1P_CHECKFORSENSORLESMODEIXXX : BOOL
VAR_INPUT
	WMCTRLMODE : WORD;
END_VAR
END_FUNCTION

(* ---- L_MC1P_CODENUMBERTOPARAMETER.pou ---- *)
FUNCTION L_MC1P_CODENUMBERTOPARAMETER : DINT
VAR_INPUT
	DWCODENUMBER : DWORD;
	USISUBINDEX : USINT;
	UIBYTELENGTH : UINT;
END_VAR
END_FUNCTION

(* ---- L_MC1P_CODENUMBERTOPARAMETER2.pou ---- *)
FUNCTION L_MC1P_CODENUMBERTOPARAMETER2 : DINT
VAR_INPUT
	DWCODENUMBER : DWORD;
	USISUBINDEX : USINT;
	UIBYTELENGTH : UINT;
	XUNSIGNED : BOOL := FALSE;
END_VAR
END_FUNCTION

(* ---- L_MC1P_CONVERTPOSTOMODULOPOS.pou ---- *)
FUNCTION L_MC1P_CONVERTPOSTOMODULOPOS : LREAL
VAR_INPUT
	LRPOS : LREAL;
	LRPERIOD : LREAL;
END_VAR
END_FUNCTION

(* ---- L_MC1P_CONVERTPOSTOMODULOPOSEXTENDED.pou ---- *)
FUNCTION L_MC1P_CONVERTPOSTOMODULOPOSEXTENDED : LREAL
VAR_INPUT
	LRPOS : LREAL;
	LRPERIOD : LREAL;
END_VAR
END_FUNCTION

(* ---- L_MC1P_CONVERTPOSTOMODULOPOSFMOD.pou ---- *)
FUNCTION L_MC1P_CONVERTPOSTOMODULOPOSFMOD : LREAL
VAR_INPUT
	LRPOS : LREAL;
	LRPERIOD : LREAL;
END_VAR
END_FUNCTION

(* ---- L_MC1P_DIV.pou ---- *)
FUNCTION L_MC1P_DIV : LREAL
VAR_INPUT
	A : LREAL;
	B : LREAL;
END_VAR
END_FUNCTION

(* ---- L_MC1P_FINDDRIVECONNECTORFROMENCODER.pou ---- *)
FUNCTION L_MC1P_FINDDRIVECONNECTORFROMENCODER : POINTER TO IoConfigConnector
VAR_INPUT
	PCONNECTOR : POINTER TO IoConfigConnector;
END_VAR
END_FUNCTION

(* ---- L_MC1P_FINDOWNSLICEPOSITIONS131.pou ---- *)
FUNCTION L_MC1P_FINDOWNSLICEPOSITIONS131 : BOOL
VAR_INPUT
	M_PCONNECTOR : POINTER TO IoConfigConnector;
END_VAR
VAR_OUTPUT
	WSLICEPOSITION : WORD;
END_VAR
END_FUNCTION

(* ---- L_MC1P_FINDPDODATAINCONNECTOR.pou ---- *)
FUNCTION L_MC1P_FINDPDODATAINCONNECTOR : POINTER TO BYTE
VAR_INPUT
	PCONNECTOR : POINTER TO IoConfigConnector;
	UIINDEX : WORD;
	USISUBINDEX : USINT;
	XWRITEACCESS : BOOL;
END_VAR
VAR_OUTPUT
	USISIZE : USINT;
END_VAR
END_FUNCTION

(* ---- L_MC1P_GENTIMESTAMPSIMU.pou ---- *)
FUNCTION L_MC1P_GENTIMESTAMPSIMU : WORD
VAR_IN_OUT
	AXIS : AXIS_REF;
END_VAR
END_FUNCTION

(* ---- L_MC1P_GETDIGINPUTSFROMDRIVE.pou ---- *)
FUNCTION L_MC1P_GETDIGINPUTSFROMDRIVE : DWORD
VAR_IN_OUT
	AXIS : AXIS_REF;
END_VAR
END_FUNCTION

(* ---- L_MC1P_GETINSTANCENAME.pou ---- *)
FUNCTION L_MC1P_GETINSTANCENAME : STRING(L_MC1P_Constants.gc_wInstanceNchar)
VAR_INPUT
	SSTR : STRING(L_MC1P_Constants.gc_wInstanceNchar);
END_VAR
END_FUNCTION

(* ---- L_MC1P_GETIOMGRCONFIGCONNECTORLIST.pou ---- *)
FUNCTION L_MC1P_GETIOMGRCONFIGCONNECTORLIST : SysTypes.RTS_IEC_RESULT
VAR_INPUT
	PPCONNECTORLIST : POINTER TO POINTER TO IoConfigConnector;
	PNCOUNT : POINTER TO DINT;
END_VAR
END_FUNCTION

(* ---- L_MC1P_GETIOMGRCONFIGFINDCONNETOR.pou ---- *)
FUNCTION L_MC1P_GETIOMGRCONFIGFINDCONNETOR : POINTER TO IoConfigConnector
VAR_INPUT
	PCONNECTOR : POINTER TO IoConfigConnector;
END_VAR
VAR_OUTPUT
	NCOUNT : DINT := 0;
END_VAR
END_FUNCTION

(* ---- L_MC1P_GETIOMGRCONFIGFIRSTCHILD.pou ---- *)
FUNCTION L_MC1P_GETIOMGRCONFIGFIRSTCHILD : POINTER TO IoConfigConnector
VAR_INPUT
	PIOCONNECTORLIST : POINTER TO IoConfigConnector;
	PNCOUNT : POINTER TO DINT;
	PFATHER : POINTER TO IoConfigConnector;
END_VAR
END_FUNCTION

(* ---- L_MC1P_GETIOMGRCONFIGNEXTCHILD.pou ---- *)
FUNCTION L_MC1P_GETIOMGRCONFIGNEXTCHILD : POINTER TO IoConfigConnector
VAR_INPUT
	PIOCONNECTORLIST : POINTER TO IoConfigConnector;
	PNCOUNT : POINTER TO DINT;
	PFATHER : POINTER TO IoConfigConnector;
END_VAR
END_FUNCTION

(* ---- L_MC1P_GETIOMGRCONFIGPARAMETER.pou ---- *)
FUNCTION L_MC1P_GETIOMGRCONFIGPARAMETER : POINTER TO IoConfigParameter
VAR_INPUT
	PCONNECTOR : POINTER TO IoConfigConnector;
	DWPARAMETERID : DWORD;
END_VAR
END_FUNCTION

(* ---- L_MC1P_GETIOMGRCONFIGPARAMETERVALUEBYTE.pou ---- *)
FUNCTION L_MC1P_GETIOMGRCONFIGPARAMETERVALUEBYTE : BYTE
VAR_INPUT
	PPARAMETER : POINTER TO IoConfigParameter;
	PRESULT : POINTER TO UDINT;
END_VAR
END_FUNCTION

(* ---- L_MC1P_GETIOMGRCONFIGPARAMETERVALUEDWORD.pou ---- *)
FUNCTION L_MC1P_GETIOMGRCONFIGPARAMETERVALUEDWORD : DWORD
VAR_INPUT
	PPARAMETER : POINTER TO IoConfigParameter;
	PRESULT : POINTER TO UDINT;
END_VAR
END_FUNCTION

(* ---- L_MC1P_GETIOMGRCONFIGPARAMETERVALUEWORD.pou ---- *)
FUNCTION L_MC1P_GETIOMGRCONFIGPARAMETERVALUEWORD : WORD
VAR_INPUT
	PPARAMETER : POINTER TO IoConfigParameter;
	PRESULT : POINTER TO UDINT;
END_VAR
END_FUNCTION

(* ---- L_MC1P_GETRATEDTORQUEAXIS.pou ---- *)
FUNCTION L_MC1P_GETRATEDTORQUEAXIS : LREAL
VAR_IN_OUT
	AXIS : AXIS_REF;
END_VAR
END_FUNCTION

(* ---- L_MC1P_GETRATEDVELOCITYAXIS.pou ---- *)
FUNCTION L_MC1P_GETRATEDVELOCITYAXIS : LREAL
VAR_IN_OUT
	AXIS : AXIS_REF;
END_VAR
END_FUNCTION

(* ---- L_MC1P_GETTASKCYCLE.pou ---- *)
FUNCTION L_MC1P_GETTASKCYCLE : LREAL
END_FUNCTION

(* ---- L_MC1P_HLPABSDINT.pou ---- *)
FUNCTION L_MC1P_HLPABSDINT : DINT
VAR_INPUT
	DIVAR : DINT;
END_VAR
END_FUNCTION

(* ---- L_MC1P_HLPCALCPOLY5THORDERSCALED.pou ---- *)
FUNCTION L_MC1P_HLPCALCPOLY5THORDERSCALED : LREAL
VAR_OUTPUT
	LRYPOSSCALED : LREAL;
END_VAR
VAR_IN_OUT
	LRXPOSSCALED : LREAL;
	ALRKOEF : ARRAY [0..5] OF LREAL;
END_VAR
END_FUNCTION

(* ---- L_MC1P_HLPCHECKDIRECTION.pou ---- *)
FUNCTION L_MC1P_HLPCHECKDIRECTION : INT
VAR_IN_OUT
	LRPOSFIFOX : ARRAY [1..20] OF LREAL;
	LRLEN : LREAL;
END_VAR
END_FUNCTION

(* ---- L_MC1P_HLPDELTAVELTIMEEXTENDED.pou ---- *)
FUNCTION L_MC1P_HLPDELTAVELTIMEEXTENDED : BOOL
VAR_INPUT
	LRVELSTART : LREAL;
	LRACCSTART : LREAL;
	LRMAXACC : LREAL;
	LRMAXJERK : LREAL;
END_VAR
VAR_OUTPUT
	LRTIME : LREAL;
	LRDIST : LREAL;
END_VAR
END_FUNCTION

(* ---- L_MC1P_HLPFITCYCLELIM.pou ---- *)
FUNCTION L_MC1P_HLPFITCYCLELIM : BOOL
VAR_INPUT
	PLRPOS : POINTER TO LREAL;
	LRLEN : LREAL;
END_VAR
END_FUNCTION

(* ---- L_MC1P_HLPGEARRES.pou ---- *)
FUNCTION L_MC1P_HLPGEARRES : LREAL
VAR_INPUT
	LRINPUT : LREAL;
	LRNUM : LREAL;
	LRDEN : LREAL;
END_VAR
END_FUNCTION

(* ---- L_MC1P_HLPMODULOADD.pou ---- *)
FUNCTION L_MC1P_HLPMODULOADD : LREAL
VAR_INPUT
	LRINPUT : LREAL;
	LROFFSET : LREAL;
	LRLENGHT : LREAL;
END_VAR
END_FUNCTION

(* ---- L_MC1P_HLPMODULODIFF.pou ---- *)
FUNCTION L_MC1P_HLPMODULODIFF : LREAL
VAR_INPUT
	LRDIFF : LREAL;
	LRLEN : LREAL;
END_VAR
END_FUNCTION

(* ---- L_MC1P_HLPMODULOOFFSET.pou ---- *)
FUNCTION L_MC1P_HLPMODULOOFFSET : LREAL
VAR_INPUT
	LROFFSET : LREAL;
	LRLENGTH : LREAL;
	PLROFFSETBASE : POINTER TO LREAL;
END_VAR
END_FUNCTION

(* ---- L_MC1P_HLPMODULOSUB.pou ---- *)
FUNCTION L_MC1P_HLPMODULOSUB : LREAL
VAR_INPUT
	LRDIFF : LREAL;
	LRLEN : LREAL;
END_VAR
END_FUNCTION

(* ---- L_MC1P_HLPMODULOZEROPOS.pou ---- *)
FUNCTION L_MC1P_HLPMODULOZEROPOS : BOOL
VAR_INPUT
	PLRPOS : POINTER TO LREAL;
	LRLENINT : LREAL;
END_VAR
END_FUNCTION

(* ---- L_MC1P_HLPPOLY4RG.pou ---- *)
FUNCTION L_MC1P_HLPPOLY4RG : LREAL
VAR_INPUT
	LRX : LREAL;
END_VAR
END_FUNCTION

(* ---- L_MC1P_HLPPT1FILT.pou ---- *)
FUNCTION L_MC1P_HLPPT1FILT : LREAL
VAR_INPUT
	LRVALUE : LREAL;
	LRINPUT : LREAL;
	LRNEW_N : LREAL;
END_VAR
END_FUNCTION

(* ---- L_MC1P_HLPSIGNNE.pou ---- *)
FUNCTION L_MC1P_HLPSIGNNE : BOOL
VAR_INPUT
	A : LREAL;
	B : LREAL;
END_VAR
END_FUNCTION

(* ---- L_MC1P_INDEXTOPARAMETER.pou ---- *)
FUNCTION L_MC1P_INDEXTOPARAMETER : DINT
VAR_INPUT
	UIINDEX : UINT;
	USISUBINDEX : USINT;
	UIBYTELENGTH : UINT := 4;
END_VAR
END_FUNCTION

(* ---- L_MC1P_INDEXTOPARAMETER2.pou ---- *)
FUNCTION L_MC1P_INDEXTOPARAMETER2 : DINT
VAR_INPUT
	UIINDEX : UINT;
	USISUBINDEX : USINT;
	UIBYTELENGTH : UINT := 4;
	XUNSIGNED : BOOL := FALSE;
END_VAR
END_FUNCTION

(* ---- L_MC1P_LMDATAMANAGERINSERTDATA.pou ---- *)
FUNCTION L_MC1P_LMDATAMANAGERINSERTDATA : BOOL
VAR_INPUT
	ITFLMDATA : L_MC1P_ILMData;
END_VAR
END_FUNCTION

(* ---- L_MC1P_LREAL_TO_DINT.pou ---- *)
FUNCTION L_MC1P_LREAL_TO_DINT : DINT
VAR_INPUT
	LRVALUE : LREAL;
END_VAR
END_FUNCTION

(* ---- L_MC1P_LREAL_TO_DINT_TO_DWORD.pou ---- *)
FUNCTION L_MC1P_LREAL_TO_DINT_TO_DWORD : DWORD
VAR_INPUT
	LRVALUE : LREAL;
END_VAR
END_FUNCTION

(* ---- L_MC1P_LREAL_TO_DWORD.pou ---- *)
FUNCTION L_MC1P_LREAL_TO_DWORD : DWORD
VAR_INPUT
	LRVALUE : LREAL;
END_VAR
END_FUNCTION

(* ---- L_MC1P_LREAL_TO_INT.pou ---- *)
FUNCTION L_MC1P_LREAL_TO_INT : INT
VAR_INPUT
	LRVALUE : LREAL;
END_VAR
END_FUNCTION

(* ---- L_MC1P_LREAL_TO_INT_TO_WORD.pou ---- *)
FUNCTION L_MC1P_LREAL_TO_INT_TO_WORD : WORD
VAR_INPUT
	LRVALUE : LREAL;
END_VAR
END_FUNCTION

(* ---- L_MC1P_LREAL_TO_WORD.pou ---- *)
FUNCTION L_MC1P_LREAL_TO_WORD : WORD
VAR_INPUT
	LRVALUE : LREAL;
END_VAR
END_FUNCTION

(* ---- L_MC1P_LREQ.pou ---- *)
FUNCTION L_MC1P_LREQ : BOOL
VAR_INPUT
	LRVALUE : LREAL;
	LRTARGET : LREAL;
END_VAR
END_FUNCTION

(* ---- L_MC1P_LRGE.pou ---- *)
FUNCTION L_MC1P_LRGE : BOOL
VAR_INPUT
	LRVALUE : LREAL;
	LRTARGET : LREAL;
END_VAR
END_FUNCTION

(* ---- L_MC1P_LRGT.pou ---- *)
FUNCTION L_MC1P_LRGT : BOOL
VAR_INPUT
	LRVALUE : LREAL;
	LRTARGET : LREAL;
END_VAR
END_FUNCTION

(* ---- L_MC1P_LRLE.pou ---- *)
FUNCTION L_MC1P_LRLE : BOOL
VAR_INPUT
	LRVALUE : LREAL;
	LRTARGET : LREAL;
END_VAR
END_FUNCTION

(* ---- L_MC1P_LRLT.pou ---- *)
FUNCTION L_MC1P_LRLT : BOOL
VAR_INPUT
	LRVALUE : LREAL;
	LRTARGET : LREAL;
END_VAR
END_FUNCTION

(* ---- L_MC1P_LRNE.pou ---- *)
FUNCTION L_MC1P_LRNE : BOOL
VAR_INPUT
	LRVALUE : LREAL;
	LRTARGET : LREAL;
END_VAR
END_FUNCTION

(* ---- L_MC1P_MODULOCYCLE.pou ---- *)
FUNCTION L_MC1P_MODULOCYCLE : LREAL
VAR_INPUT
	LRPOSIN : LREAL;
	LRPOSITIONPERIOD : LREAL;
END_VAR
END_FUNCTION

(* ---- L_MC1P_POS_DINT_TO_LINT.pou ---- *)
FUNCTION L_MC1P_POS_DINT_TO_LINT : LINT
VAR_INPUT
	DIPOS : DINT;
	DIPOSOLD : DINT;
END_VAR
VAR_IN_OUT
	UPOS : L_MC1P_PosLINT;
END_VAR
END_FUNCTION

(* ---- L_MC1P_POSDIFFTOSPEEDINCIXXX.pou ---- *)
FUNCTION L_MC1P_POSDIFFTOSPEEDINCIXXX : DINT
VAR_INPUT
	DIPOSDIFF : DINT := 0;
	DWFACTOR : DWORD := 1000;
	DWINKPERREV : DWORD := 65536;
END_VAR
END_FUNCTION

(* ---- L_MC1P_SPEEDTOPOSDIFFINCIXXX.pou ---- *)
FUNCTION L_MC1P_SPEEDTOPOSDIFFINCIXXX : DINT
VAR_INPUT
	DISPEED : DINT := 0;
	DWFACTOR : DWORD := 1000;
	DWINKPERREV : DWORD := 65536;
END_VAR
VAR_IN_OUT
	DIRES : DINT;
END_VAR
END_FUNCTION

(* ---- L_MC1P_STVARIABLENAME_TO_DWORD.pou ---- *)
FUNCTION L_MC1P_STVARIABLENAME_TO_DWORD : BOOL
VAR_INPUT
	STVARIABLENAME : STRING;
END_VAR
VAR_OUTPUT
	DWOUT : DWORD;
END_VAR
END_FUNCTION

(* ---- L_MC1P_STVARIABLENAME_TO_INT.pou ---- *)
FUNCTION L_MC1P_STVARIABLENAME_TO_INT : BOOL
VAR_INPUT
	STVARIABLENAME : STRING;
END_VAR
VAR_OUTPUT
	IOUT : INT;
END_VAR
END_FUNCTION

(* ---- L_MC1P_STVARIABLENAME_TO_LREAL.pou ---- *)
FUNCTION L_MC1P_STVARIABLENAME_TO_LREAL : BOOL
VAR_INPUT
	STVARIABLENAME : STRING(255);
END_VAR
VAR_OUTPUT
	LROUT : LREAL;
END_VAR
END_FUNCTION

(* ---- L_MC1P_STVARIABLENAME_TO_REAL.pou ---- *)
FUNCTION L_MC1P_STVARIABLENAME_TO_REAL : BOOL
VAR_INPUT
	STVARIABLENAME : STRING;
END_VAR
VAR_OUTPUT
	ROUT : REAL;
END_VAR
END_FUNCTION

(* ---- L_MC1P_STVARIABLENAME_TO_WORD.pou ---- *)
FUNCTION L_MC1P_STVARIABLENAME_TO_WORD : BOOL
VAR_INPUT
	STVARIABLENAME : STRING;
END_VAR
VAR_OUTPUT
	WOUT : WORD;
END_VAR
END_FUNCTION

(* ---- L_MC1P_TRUNC_LINT.pou ---- *)
FUNCTION L_MC1P_TRUNC_LINT : LINT
VAR_INPUT
	LRIN : LREAL;
END_VAR
END_FUNCTION

(* ---- L_MC1P_USEHOMINGPOSITIONFROMAXISREF.pou ---- *)
FUNCTION L_MC1P_USEHOMINGPOSITIONFROMAXISREF : BOOL
VAR_INPUT
	XACTIVATE : BOOL;
END_VAR
VAR_IN_OUT
	AXIS : AXIS_REF;
END_VAR
END_FUNCTION

(* ---- L_MC1P_USEMANUALPARAMETERFROMAXISREF.pou ---- *)
FUNCTION L_MC1P_USEMANUALPARAMETERFROMAXISREF : BOOL
VAR_INPUT
	XACTIVATE : BOOL;
END_VAR
VAR_IN_OUT
	AXIS : AXIS_REF;
END_VAR
END_FUNCTION

(* ---- AXIS_REF.pou ---- *)
FUNCTION_BLOCK AXIS_REF EXTENDS L_DCO_AXIS_REF_BASE
VAR_INPUT
	LRVELOVERRIDE : LREAL := 1.0;
	LRACCOVERRIDE : LREAL := 1.0;
	LRJERKOVERRIDE : LREAL := 1.0;
	LRCOMMANDEDPOSITION : LREAL;
	LRCOMMANDEDVELOCITY : LREAL;
	LRCOMMANDEDACCELERATION : LREAL;
	LRSETVELOCITYLIMITHIGH : LREAL := 0;
	LRSETVELOCITYLIMITLOW : LREAL := 0;
	LRTORQUELIMHIGH : LREAL;
	LRTORQUELIMLOW : LREAL;
	LRTORQUELIMAUX : LREAL;
	SITORQUELIMDIR : SINT;
	XDELETETORQUELIM : BOOL;
	XSETTORQUELIMAUX : BOOL;
	XTORQUELIMHIGHFROMAPP : BOOL;
	XTORQUELIMLOWFROMAPP : BOOL;
	ITORQUELIMHIGHPCT : INT := 2000;
	ITORQUELIMLOWPCT : INT := 2000;
	EDIRECTION : MC_DIRECTION;
	XDRIVEENABLE : BOOL;
	XERRORRESET : BOOL;
	LRREFOFFSET : LREAL;
	LRREFOFFSETACT : LREAL;
	XENABLEPOSITIVE : BOOL := TRUE;
	XENABLENEGATIVE : BOOL := TRUE;
	LRSETSUPERACC : LREAL;
	LRSETSUPERVEL : LREAL;
	LRSETSUPERPOS : LREAL;
	LRSETMOVEACC : LREAL;
	LRSETMOVEVEL : LREAL;
	LRSETMOVEPOS : LREAL;
	XBUFCMDDONE : BOOL;
	XBUFRESTART : BOOL;
	LRPROFILESPEEDFIRST : LREAL;
	LRPROFILETARGETSPEED : LREAL;
	DWBUFFERCMD : __XWORD;
	XDISABLEERRORLOGGING : BOOL;
	XMOVEFUNBUSY : BOOL;
	XSUPERFUNBUSY : BOOL;
	LRCOMMANDEDPOSABSOLUT : LREAL;
	XRESETFOLLOWINGERROR : BOOL;
	XSETAXISQSP : BOOL;
	XSETDRIVEQSP : BOOL;
	EAXISSTATE : L_MC1P_AXIS_STATE := 2;
	LRSETPOSITION : LREAL := 0.0;
	LRSETVELOCITY : LREAL := 0.0;
	LRSETACCELERATION : LREAL := 0.0;
	LRSETTORQUE : LREAL := 0.0;
	LRVLTARGETVEL : LREAL := 0.0;
	LRLIMITEDVELOCITY : ARRAY [1..4] OF LREAL;
	LRLIMITEDDECTIME : ARRAY [1..4] OF LREAL;
	LRRESETSLSOFFSETVELOCITY : LREAL;
	DWLIMITERCONTROLACT : DWORD;
	SCSTOPAXISBYAPPL : L_MC1P_StopOperation;
	XSTAYINLASTSTATEREQUEST : BOOL;
	XMOVELASTSETPOSREQUEST : BOOL;
	LRSETVELMOVELASTSETPOS : LREAL;
	LRSETACCMOVELASTSETPOS : LREAL;
	LRSETDECMOVELASTSETPOS : LREAL;
	LRSETJERKMOVELASTSETPOS : LREAL;
	EDIRECTIONMOVELASTSETPOS : MC_DIRECTION;
	EDIRECTIONACTPROFILE : MC_DIRECTION;
	WAXISCONTROL : WORD := 0;
	XALLOWCHANGEOFCINHPAR : BOOL := FALSE;
	LRMOVEVELOFFSETVEL : LREAL;
	EOPTIMIZEDPROFILECALCULATIONMODE : UINT := 1;
	XENABLECOMPOFFSET : BOOL := TRUE;
	XCOMPQSPACCOFFSET : BOOL := FALSE;
	WMODECOMP : WORD;
END_VAR
VAR_OUTPUT
	EDEVICE : L_MC1P_DriveType := 0;
	WAXISSTATUS : DWORD := 0;
	EACTIVEERRORID : WORD := 0;
	LRACTPOSITION : LREAL := 0.0;
	LRACTVELOCITY : LREAL := 0.0;
	LRACTACCELERATION : LREAL := 0.0;
	LRACTTORQUE : LREAL := 0.0;
	LRSETTORQUETODRIVE : LREAL := 0;
	LRACTFOLLOWINGERROR : LREAL := 0.0;
	LRMAXFOLLOWINGERROR : LREAL := 0.0;
	XVIRTUAL : BOOL;
	XAXISAVAILABLE : BOOL;
	EACTDIRECTION : MC_DIRECTION;
	LRDIRECTIONHYSTERESISPOS : LREAL;
	LRDIRECTIONHYSTERESISTOL : LREAL := 1E-06;
	XDRIVEENABLED : BOOL;
	XERROR : BOOL;
	XWARNING : BOOL;
	XDRIVEERROR : BOOL;
	XDRIVEWARNING : BOOL;
	DWDRIVEERRORID : DWORD;
	XHOMEPOSAVAILABLE : BOOL;
	XSWLIMITENABLED : BOOL;
	XSWLIMITPOS : BOOL;
	XSWLIMITNEG : BOOL;
	XHWLIMITPOS : BOOL;
	XHWLIMITNEG : BOOL;
	XSPEEDEQZERO : BOOL;
	XINPOSITION : BOOL;
	LRTASKCYCLE : LREAL := 0.001;
	LRINVTASKCYCLE : LREAL := 1000.0;
	LRSWLIMITPOS : LREAL := 0.0;
	LRSWLIMITNEG : LREAL := 0.0;
	LRLASTSETPOSITION : LREAL;
	LRLASTTARGETPOSITION : LREAL;
	XSTANDSTILLSETVELOCITY : BOOL;
	XSTANDSTILLACTVELOCITY : BOOL;
	XSTOACTIVE : BOOL;
	XVOLTAGEENABLED : BOOL;
	XAXISREADYTOSWITCHON : BOOL;
	XAXISREADYFORMOTION : BOOL;
	SCPAR : L_MC1P_ParAccess;
END_VAR
VAR
	AXISTASKIDX : INT;
	XMCFEATUREUSED : BOOL := FALSE;
	AXISVALUESTORE : L_MC1P_AxisValueStore;
	DWAXISCONFIGSETTINGS : DWORD;
	XSETVALUESAVAILABLE : BOOL;
	BYSETVALUESVALID : BYTE;
	DWTASKYCLE_US : DWORD := 1000;
	XSUSPENDFOLLOWINGERRORINT : BOOL;
	XSUSPENDFOLLOWINGERROREXT : BOOL;
	LRMAXVELOCITYAPPLOLD : LREAL;
	LRMAXACCELERATIONAPPLOLD : LREAL;
	LRMAXJERKAPPLOLD : LREAL;
	LRSWLIMITPOSOLD : LREAL;
	LRSWLIMITNEGOLD : LREAL;
	XENABLEPOSOLD : BOOL;
	XENABLENEGOLD : BOOL;
	DWLIMITERCONTROLOLD : DWORD;
	LRLIMITEDVELOCITYOLD : ARRAY [1..4] OF LREAL;
	LRLIMITEDDECTIMEOLD : ARRAY [1..4] OF LREAL;
	LRLIMITEDJERKOLD : ARRAY [1..4] OF LREAL;
	ELIMITERSTOPREACTION : L_IE1P_SeverityLevel := L_IE1P_SeverityLevel.WARNING;
	XSWLIMITDISABLE : BOOL := FALSE;
	XSWLIMITPOSNEU : BOOL;
	XSWLIMITPOSISTAN : BOOL;
	XSWLIMITNEGNEU : BOOL;
	XSWLIMITNEGISTAN : BOOL;
	PBYCOUPLEDMASTERAXIS : POINTER TO BYTE;
	PBYCOUPLEDPHASINGMASTERAXIS : POINTER TO BYTE;
	LRPHASESHIFTPOS : LREAL;
	LRPHASESHIFTVEL : LREAL;
	LRPHASESHIFTACC : LREAL;
	LRPHASESHIFTPOSOLD : LREAL;
	LRPHASESHIFTVELOLD : LREAL;
	LRPHASESHIFTACCOLD : LREAL;
	XSETPHASESHIFTVALUES : BOOL;
	ETRAVERSINGRANGEACT : L_MC1P_TraversingRange := 0;
	LRCYCLELENGTHACT : LREAL := 360.0;
	XENABLEHWLIMITPOS : BOOL := TRUE;
	XENABLEHWLIMITNEG : BOOL := TRUE;
	XHWSIGNALNEG : BOOL := FALSE;
	XHWSIGNALPOS : BOOL := FALSE;
	BHWENSCHPOSNEU : BOOL := TRUE;
	BNOTIFYERRORHWLIMITPOSISTAN : BOOL;
	BHWENSCHNEGNEU : BOOL := TRUE;
	BNOTIFYERRORHWLIMITNEGISTAN : BOOL;
	XAXISISHOMESOURCE : BOOL;
	XHOMEPOSAVAILABLEDRIVE : BOOL;
	SCHOMEPARAMETER : L_MC1P_HomeParameter;
	LRHOMEPOSITION : LREAL;
	XPOSCTRL : BOOL;
	XTPSUPPORTED : BOOL := FALSE;
	XTPWITHTIMESTAMP : BOOL := FALSE;
	SNTPMAXCHANNEL : SINT;
	PG : L_MC1P_PosProfiler := STRUCT(wCalcProfileMode := 1);
	ITFPG_MOVEACTIVE : L_MC1P_IPosProfilerActive;
	PG_MOVE : L_MC1P_PosProfiler := STRUCT(wCalcProfileMode := 1);
	ITFPG_SUPERACTIVE : L_MC1P_IPosProfilerActive;
	PG_SUPER : L_MC1P_PosProfiler := STRUCT(wCalcProfileMode := 1);
	PG_DUMMY : L_MC1P_PosProfiler := STRUCT(wCalcProfileMode := 1);
	SCPARAMSTOP : L_MC1P_ProfileParameter;
	XCTRLMODECHANGEREQ : BOOL;
	LRCTRLMODECHANGEREQACTVEL : LREAL;
	PFBMOVEBASIC : POINTER TO L_MC1P_MoveBasic;
	PFBMOVEBASICSUPER : POINTER TO L_MC1P_MoveBasic;
	XRESTARTPOSITIONING : BOOL;
	LRSETPOSITIONOLD : LREAL;
	LRSETVELOCITYOLD : LREAL;
	LRSETACCELERATIONOLD : LREAL;
	WACTFUNID : WORD := 0;
	WACTSUPERFUNID : WORD := 0;
	WACTPHASEFUNID : WORD := 0;
	PSERRORINST : POINTER TO STRING;
	SERRORINST : STRING;
	ERRORMANAGER : L_IE1P_ErrorManager;
	ERRORRESETOCCUREDTIMEWITHOUTLEM : SYSTIME;
	ASCERRORINFO : REFERENCE TO ARRAY [0..7] OF L_IE1P_ErrorInformation;
	ASCWARNINGINFO : REFERENCE TO ARRAY [0..7] OF L_IE1P_ErrorInformation;
	WINITSTATE : WORD;
	PAPPLICATION : POINTER TO APPLICATION;
	ATPDATA : ARRAY [1..4] OF L_MC1P_TPData;
	ATPDATASAVE : L_MC1P_TPData;
	XHOMINGSUPPORTED : BOOL;
	EAXISSTATEOLD : L_MC1P_AXIS_STATE := L_MC1P_AXIS_STATE.Disabled;
	ECONTROLMODE : L_MC1P_ControlMode := L_MC1P_ControlMode.PosCtrlDrive;
	ECONTROLMODEDEFAULT : L_MC1P_ControlMode := L_MC1P_ControlMode.PosCtrlDrive;
	ECONTROLMODEDEFAULTINT : L_MC1P_ControlMode := L_MC1P_ControlMode.PosCtrlDrive;
	POSCTRLDRIVEAVAILABLE : L_IE1P_Error;
	POSCTRLPLCAVAILABLE : L_IE1P_Error;
	SPEEDCTRLDRIVEAVAILABLE : L_IE1P_Error;
	TORQUECTRLDRIVE : L_IE1P_Error;
	XDRIVEENABLEOLD : BOOL;
	XLOCKEDFORSINGLEMOTION : BOOL := FALSE;
	XHOMEABSSWITCH : BOOL;
	XHOMEABSSWITCHOVERWRITEACTIVE : BOOL;
	XRAMPTOSTANDSTILL : BOOL;
	XRAMPTOSTANDSTILLDONE : BOOL;
	XRAMPTOSTANDSTILLACTIVE : BOOL;
	XRAMPDOWNINSERVICESTATE : BOOL;
	XDRIVEENABLEDOLD : BOOL;
	XDRIVEENABLEDREAL : BOOL;
	XDRIVEENABLEDREALOLD : BOOL;
	LRFOLLOWINGERRORINT : LREAL;
	XSUPPORTBRAKE : BOOL := FALSE;
	XSUPPORTDCBRAKE : BOOL := FALSE;
	XUSEASVIRTUALEXT : BOOL := FALSE;
	XUSEASVIRTUALEXTACT : BOOL := FALSE;
	LRSETSUPERACCOLD : LREAL;
	LRSETSUPERVELOLD : LREAL;
	LRSETSUPERPOSOLD : LREAL;
	ITFPARA : L_MC1P_IPara;
	XFASTSTOPDONE : BOOL;
	XFASTSTOPDONESAVE : BOOL;
	XSETFASTSTOPINT : BOOL;
	XERRRORSTOPACTIVE : BOOL;
	XERRRORSTOPDONE : BOOL;
	XSETAXISQSPACTIVE : BOOL;
	XRAMPQSPSTARTCALLEDFROMAPP : BOOL;
	XDRIVEQSPACTIVE : BOOL;
	XDRIVEFAULTREACTIONACTIVE : BOOL;
	XDRIVEQSPACTIVEOLD : BOOL;
	XDRIVEQSPSET : BOOL;
	XSTOPINDISABLEDALLOWED : BOOL;
	XSETDRIVEFAILQSP : BOOL;
	XSETDRIVEFAILCINH : BOOL;
	XDRIVEQSPDONE : BOOL;
	XDRIVEQSPDONESAVE : BOOL;
	ESTOPTYPE : WORD;
	POW : L_MC1P_Power_Internal;
	XOBERVERESWITCHONTIME : BOOL := TRUE;
	FBBASE : L_MC1P_Template_ForAxis;
	ABC : L_MC1P_AxisBasicControl_Internal;
	ABCDATA : L_MC1P_AxisBasicControlInstanceData;
	ITFENCODER : L_MC1P_IEncoderInterface;
	ITFENCODERHANDLER : L_MC1P_IEncoderInterface;
	LRSETTORQUEFROMAXESGROUP : LREAL := 0;
	EPRECONTROLMODE : L_MC1P_PreControlMode := L_MC1P_PreControlMode.Automatic;
	GUID : L_MC1P_AxisGUID;
	LRTORQUEPRECTRL : LREAL;
	LRTORQUESET : LREAL;
	XMOVEFUNBUSYOLD : BOOL;
	XMOVEFUNBUSYOLDOLD : BOOL;
	DWIODRVDEVICEID : DWORD;
	WIODRVDEVICETYPE : WORD;
	EDEVICEORIGIN : L_MC1P_DriveType := L_MC1P_DriveType.Virtual;
	EDEVICECLASS : L_MC1P_DeviceClass := L_MC1P_DeviceClass.VirtualAxis;
	DWTARGETID : DWORD := 0;
	XCTRLFIRMWARECHECKPASSED : BOOL := FALSE;
	XENABLELOGENTRY : BOOL := 1;
	ETRAVERSINGRANGE : L_MC1P_TraversingRange := 1;
	LRCYCLELENGTH : LREAL := 360.0;
	LRINVCYCLELENGTH : LREAL := (1.0 / 360.0);
	LRDEFAULTVELOCITY : LREAL := 0.0;
	LRDEFAULTACCELERATION : LREAL := 0.0;
	LRDEFAULTJERK : LREAL := 0.0;
	LRMAXVELOCITYAPPL : LREAL := 0.0;
	LRMAXACCELERATIONAPPL : LREAL := 0.0;
	LRMAXJERKAPPL : LREAL := 0.0;
	XENABLESWLIMIT : BOOL := 0;
	WBEHAVEONSWLIMIT : WORD := 1;
	LRDECERRORSTOP : LREAL := 3600.0;
	LRJERKERRORSTOP : LREAL := 0.0;
	XREAKTONMCFBERROR : BOOL := 1;
	LRWINDOWSTANDSTILL : LREAL := 0.0;
	LRWINDOWVELOCITYCONST : LREAL := 0.0;
	LRWINDOWTARGETREACHED : LREAL := 0.0;
	LRWINDOWTARGETREACHEDTIME : LREAL := 0.0;
	LRMODPOSTOLERANCE : LREAL := 0.0;
	XSETVALUEMONITORING : BOOL := 0;
	EPARAMETERINDEX : WORD := 101;
	DWPARABASEINDEX : DWORD;
	PPARA2 : L_SSYP.L_SSYP_EVTPARAM_CmpLenzeIPCSystemSoftPLCParaChanged;
	HEVENTPARWRITE : SysTypes.RTS_IEC_HANDLE;
	HINTERFACEPARWRITE : SysTypes.RTS_IEC_HANDLE;
	HEVENTDOWNLOADDONE : SysTypes.RTS_IEC_HANDLE;
	HINTERFACEDOWNLOADDONE : SysTypes.RTS_IEC_HANDLE;
	HEVENTRESETDONE : SysTypes.RTS_IEC_HANDLE;
	HINTERFACERESETDONE : SysTypes.RTS_IEC_HANDLE;
	ITFCALLBACK : CmpEventMgr.ICmpEventCallback;
	DWEVENTCOUNTER : DWORD;
	WENABLEDRIVEBLOCKEDBYOBJECTTRANSFER : WORD := 0;
	XUSEDBYAXESGROUP : BOOL;
	PUSEDAXESGROUP : POINTER TO BYTE;
	DWEVTINITCOUNT : DWORD;
	XNEWHOMEPOSLOADED : BOOL;
	DWSETPOSITIONCALLCYCLE : DWORD;
	XSETPOSITIONCALLCYCLEVALID : BOOL;
	AITFFILTER : ARRAY [1..c_MaxFilterInt] OF L_MC1P_ISetvalueManipulationInterface;
	XENABLEFILTER : BOOL;
	XFILTERAVAILABLE : BOOL;
	XIGNORFILTERINSTOP : BOOL := TRUE;
	XIGNORFILTERINSTOPITF : BOOL;
	XUSEFILTERVALUESFORSYNC : BOOL := FALSE;
	LRSETPOSITIONFILT : LREAL;
	LRSETVELOCITYFILT : LREAL;
	LRSETACCELERATIONFILT : LREAL;
	LRSETTORQUEFILT : LREAL;
	LRSETVALUEFILTERPOSDEVIATION : LREAL;
	XINTARGETSETVALUEFILTER : BOOL;
	XSUSPENDSETVALUEFILTERCALL : BOOL := FALSE;
	LRSETPOSITIONFILTOLD : LREAL;
	LRSETVELOCITYFILTOLD : LREAL;
	LRSETACCELERATIONFILTOLD : LREAL;
	LRSETTORQUEFILTOLD : LREAL;
	LRSETPOSROUNDSFILTOLD : LREAL;
	AITFCOMPENSATION : ARRAY [1..c_MaxFilterInt] OF L_MC1P_ICompensationInterface;
	LRCOMPENSATIONOFFSETPOS : LREAL;
	LRCOMPENSATIONOFFSETVEL : LREAL;
	LRCOMPENSATIONOFFSETACC : LREAL;
	LRACTPOSITIONUNFILTERED : LREAL;
	LRINTARGETPOS : LREAL;
	LRACTTIMETARGETREACHED : LREAL;
	XSETVALUEINTARGET : BOOL;
	XUSEACYCLIC : BOOL := FALSE;
	XFORCEACYCLICMODE : BOOL := FALSE;
	WAXISMODE : WORD := 1;
	WAXISMODEOLD : WORD := 255;
	LRTRANSMITCYCLESACTPOS : LREAL := 0.0;
	LRTRANSMITCYCLESSETPOS : LREAL := 1.0;
	XCONNECTORDISABLEDBYPROJECT : BOOL;
	XCONNECTORDISABLED : BOOL;
	XAXISDETECTIONBUSY : BOOL;
	XAXISDETECTED : BOOL;
	XCONFIGDONE : BOOL;
	XBASICINIT : BOOL := TRUE;
	XAXISCONNECTBUSY : BOOL;
	XAXISCONNECTDONE : BOOL;
	XPDOINTERFACEDISABLED : BOOL;
	XDRIVETESTMODEACTIVE : BOOL;
	LRACTPOSROUNDS : LREAL;
	LRSETPOSROUNDS : LREAL;
	LRSETPOSROUNDSFILT : LREAL;
	LRSETPOSROUNDSLAST : LREAL;
	LRTARGETPOSROUNDS : LREAL;
	XTARGETPOSVALID : BOOL;
	XTARGETPOSFROMMOVEREL : BOOL;
	LISETPOSCYCLE : LINT;
	LISETPOSCYCLERES : UDINT;
	XSETPOSCYCLEZERO : BOOL;
	XRECOVERLASTSETPOS_RAMP : BOOL := FALSE;
	XRECOVERLASTSETPOS_POSCTRL : BOOL := TRUE;
	XVFCMODE : BOOL := FALSE;
	XRECOVERYPOSVALID : BOOL;
	XMOVELASTSETPOS : BOOL;
	LRRECOVERYWINDOWPOS : LREAL;
	LRRECOVERYWINDOWNEG : LREAL;
	LRRECOVERYPOSITION : LREAL;
	LRRECOVERYVEL : LREAL := 360;
	LRRECOVERYACC : LREAL := 3600;
	LRRECOVERYDEC : LREAL := 3600;
	LRRECOVERYJERK : LREAL := 0;
	XSLSACTIVE : BOOL;
	XSLSACTIVEOLD : BOOL;
	XSLIREQUESTACTIVE : BOOL;
	XSWLIMITSACTIVE : BOOL;
	LRSLIDISTANCE : LREAL := 360;
	LRSLSVELOCITY : LREAL;
	LRSLSVELOCITYOLD : LREAL;
	LRSLSDECELERATION : LREAL;
	LRSLSDECELERATION2 : LREAL;
	LRSLSDECELERATIONOLD : LREAL;
	LRSLSJERK : LREAL;
	XSLSCHANGES : BOOL;
	XSLSNEWACTIVEDECELERATION : BOOL;
	WSLSWARNING : WORD;
	XLIMITERENABLEPOSITIVE : BOOL := TRUE;
	XLIMITERENABLENEGATIVE : BOOL := TRUE;
	XLIMITERENABLED : BOOL;
	XLIMITATIONSLSACTIVE : BOOL;
	XLIMITATIONACTIVE : BOOL;
	LRSLSDECTIME : LREAL := 100;
	LRSLSDECTIMEOLD : LREAL := 100;
	WSAFESTOPCONTROLWORD : WORD;
	WSAFESTOPCONTROLWORDOLD : WORD;
	READPARAMETER : L_DCO_ReadDriveParameter;
	WRITEPARAMETER : L_DCO_WriteDriveParameter;
	DWACTUALSPEEDCONTROLLERLIMIT : DWORD;
	XLIMITSPEEDCONTROLLERSLS : BOOL;
	DWDISABLESAFETYINTERFACE : DWORD;
	DWREQUESTSAFETYINTERFACE : DWORD;
	XFOLLOWERSLS : BOOL;
	LRSLSTIMER : LREAL;
	LRSLSTIMERTEMP : LREAL;
	XSLSACTIVATED : BOOL := FALSE;
	XSETSTOPBYDIRECTIONACTIVE : BOOL;
	XSETSTOPBYLIMITERACTIVE : BOOL;
	XSETSTOPCINHBYLIMITERACTIVE : BOOL;
	XSLSVELOCITYACTIVE : BOOL;
	XSLSDECTIMEACTIVE : BOOL;
	XSLSWARNINGACTIVE : BOOL;
	ETYPEFUNCTIONACT : L_MC1P_TypeFunction := L_MC1P_TypeFunction.Type_Any;
	SCSTOPBYERROR : L_MC1P_StopOperation;
	SCSTOPBYAXESGROUP : L_MC1P_StopOperation;
	DWAXISERRORITFID : DWORD := 0;
	ICMODE : WORD;
	ICMODEOLD : WORD;
	DWIC : DWORD;
	DWICOLD : DWORD;
	XINTERNALCONTROLMODEACTIVE : BOOL;
	XINTERNALCONTROLMODEACTIVEOLD : BOOL;
	XREFDUMMY : BOOL;
	LRREFDUMMY : LREAL;
	RREFDUMMY : REAL;
	WREFDUMMY : WORD;
	IREFDUMMY : INT;
	DWREFDUMMY : DWORD;
	DIREFDUMMY : DINT;
	LWREFDUMMY : LWORD;
	LIREFDUMMY : LINT;
	SREFDUMMY : STRING;
	USIREFDUMMY : USINT;
	BYREFDUMMY : BYTE;
	UIREFDUMMY : UINT;
	UDIREFDUMMY : UDINT;
	ULIREFDUMMY : ULINT;
	DWCALLCYCLE : DWORD;
	DWCALLCYCLE_US : DWORD;
	DWTPDELAYACTPOS : DWORD := 0;
	DWACTDCTIME : DWORD;
	DWACTDCTIME_CYCLE : DWORD;
	PDWABSOLUTECOUNTER : POINTER TO DWORD;
	XGLOBALTIMESTAMPSUPPORTED : BOOL;
	HMOTIONTASK : SysTypes.RTS_IEC_HANDLE := 0;
	WACTPOSIDX : WORD;
	ADWACTTIMESTAMPS : ARRAY [0..15] OF DWORD;
	ALRACTPOSITION : ARRAY [0..15] OF LREAL;
	ALRACTPOSITIONUNFILTERED : ARRAY [0..15] OF LREAL;
	ALRACTPOSROUNDS : ARRAY [0..15] OF LREAL;
	ALRTPPOSOFFSET : ARRAY [0..15] OF LREAL;
	HEVENTRESETOCCURED : SysTypes.RTS_IEC_HANDLE := SysTypes.RTS_INVALID_HANDLE;
	HINTERFACERESETOCCURED : SysTypes.RTS_IEC_HANDLE := SysTypes.RTS_INVALID_HANDLE;
	XGENERRORREAKTINDEVICE : BOOL;
	XFORWARDERRORSASWARNINGS : BOOL;
	WEVTCOUNT_SETERRORREACTION : WORD;
	WEVTCOUNT_UPDATEACTIVEERROR : WORD;
	WEVTCOUNT_RESETOCCURED : WORD;
	XINTERNALERRORRESET : BOOL;
	XINTERNALERRORRESETFROMLEM : BOOL;
	WHANDLINGLEM : WORD := 0;
	XERRORRESETREQUESTSEND : BOOL;
	WERRORRESETREQUESTSEND : WORD := 0;
	RESETINTERNAL : L_MC1P_Reset_Internal;
	SCRESETINPUT : L_MC1P_ResetInput;
	SCRESETOUTPUT : L_MC1P_ResetOutput;
	DWACTSTATEDETERMINEEVENT : DWORD;
	SEVERITYCMDEXT : USINT;
	EERRORREACTIONCMDEXT : L_IE1P_SeverityLevel := L_IE1P_SeverityLevel.NO_RESPONSE;
	DWERRORINFOEXT : DWORD;
	XEXTERROR : BOOL;
	MYSYSTEMSEVERITY : USINT;
	XJOGGINGACTIVE : BOOL;
	LRJOGGINGSETVEL : LREAL := 360.0;
	LRJOGGINGSETACC : LREAL := 360.0;
	LRJOGGINGSETDEC : LREAL := 1440.0;
	LRJOGGINGSETJERK : LREAL := 0.0;
	XJOGUSEAXISPAR : BOOL := FALSE;
	XHOMEPOSUSEAXISPAR : BOOL := FALSE;
	XUSEFASTSTOPBEHAVIOUR : BOOL := TRUE;
	XFIRSTBASEINITDONE : BOOL := FALSE;
	EHWLIMITERRORREACTION : USINT := 19;
	ESWLIMITERRORREACTION : USINT := 19;
	ELIMITPROFILEERRORREACTION : USINT := 2;
	ECINHERRORREACTION : USINT := 19;
	LRREFROUNDS : LREAL;
	XMOVELASTSETPOSACTIVE : BOOL;
	XSTAYINLASTSTATEACTIVE : BOOL;
	XABORTSTAYINLASTSTATEREQUEST : BOOL;
	XCINHACTIVE : BOOL;
	XCINHACTIVEOLD : BOOL;
	XSTOACTIVEOLD : BOOL;
	XSETPOSINSIDEWINDOW : BOOL;
	XSTAYINLASTSTATEACTIVEOLD : BOOL;
	XDRIVESTATEBEFORECINH : BOOL;
	LRPOSOFFSETMOVELASTSETPOS : LREAL;
	LRVELOFFSETMOVELASTSETPOS : LREAL;
	LRACCOFFSETMOVELASTSETPOS : LREAL;
	XHALTPARAMETERSUPPORTED : BOOL;
	LRHALTDEC : LREAL := 1800;
	LRHALTJERK : LREAL := 0;
	XHALTBYABC : BOOL;
	SCTIMESTAMP : L_MC1P_TimeStamp;
	XACTIVATETIMEMEASUREMENT : BOOL;
	XISSAFETYDEVICE : BOOL;
	WINDEXINT : WORD;
	BYSUBINDEXINT : BYTE;
	BYSLSREADWRITECOUNTER : BYTE;
	XCALCMODULOASLIMITED : BOOL := FALSE;
	FBSTEADYSTATE : L_MC1P_SteadyState;
	WDEVICETYPETEMP : WORD;
	DWIODRVDEVICEIDTEMP : DWORD;
	XUSEQSPDRIVEINSTEADOFQSPAPPL : BOOL := FALSE;
	XMINJERKAVAILABLE : BOOL;
	XMINJERKAVAILABLEOLD : BOOL;
	XMINJERKACTIVE : BOOL;
	XMINJERKACTIVEOLD : BOOL;
	LRMINJERK : LREAL;
	LRMINJERKOLD : LREAL;
	LRMOVEVELOFFSETVELOLD : LREAL;
	XSETVALUESFORINTERNALSTOPAVAILABLE : BOOL;
	XSETVALUESFROMINTERNALSTOPACTIVE : BOOL;
	XOPTRAMPSFORMANUALJOG : BOOL := TRUE;
	XCHANGECINHPARNOTALLOWED : BOOL := FALSE;
	XBEHAVIOURFORVIRTUALMASTER : BOOL := FALSE;
	STOPAXISBYERRORREACTIONCOUNTER : L_IE1P_ReactionCounter;
	SCSTOPAXISBYERRORREACTION : L_MC1P_StopOperation;
	MODULEHANDLERBASE : L_IMHP_ModuleHandler := STRUCT(CompActiveDefault := FALSE, Layer := L_IMHP_Layer.Motion, CompType := L_IMHP_ComponentType.VirtualAxis);
	FB_GETDIRECTIONACTVALUES : L_MC1P_GetDirection;
	WDIRECTIONSETVALUES : WORD;
	XQSPWITHOUTREACTION : BOOL;
	XVALIDMFEFWVERSION : BOOL;
	XSETDRIVEQSPDISABLED : BOOL;
	EKINDOFMOTIONSELECTION : L_MC1P_KindOfMotion;
	EACTIVEUNIT : WORD;
	WERRORIDINITSTATE : WORD;
	ITFMANIPULATEACTVALUES : L_Mc1P_IManipulateActValues;
	XSETVELOCITYGTSLS : BOOL;
	XCLOSEBRAKEATQSPRAMPEND : BOOL;
	CRITICALSECTIONERRORENTRY : L_MC1P_CriticalSection;
	CRITICALSECTIONERRORREACTION : L_MC1P_CriticalSection;
	ITFSLAVEKIN : L_MC1P_IKinematicSlave;
	ITFMASTERKIN : L_MC1P_IKinematicMaster;
	XSELECTEDFORKINEMATIC : BOOL;
	XHOMINGDONEOWNAXIS : BOOL;
	XSUSPENDSWLIMITERRORREACTION : BOOL;
	XWRITEOUTPUTWASCALLED : BOOL := FALSE;
	XREADINPUTSWASCALLED : BOOL := FALSE;
	ITFCALLDEPENDENCYKINEMATIC : L_UBUP_ICallOrderDependency;
	DWAXISINTERNALCONTROL : DWORD;
	WINTERNALCONTROLSTATUS : WORD;
	LRICJOGDISTANCE : LREAL := 10.0;
	IICJOGOVERRIDE : INT := 100;
	XGRINDINDONEOWNAXIS : BOOL;
	XBRAKETESTDONEOWNAXIS : BOOL;
	POWIDGI : WORD;
	POWIDBT : WORD;
	ALRQSPAPPLOFFSET : ARRAY [0..2] OF LREAL;
	XCOMPPOSOFFSET : BOOL;
	XCOMPOFFSETDONE : BOOL;
	XCOMPOFFSETBUSY : BOOL;
	XEXECUTECOMPOFFSET : BOOL;
	XCOMPPOSOFFESTALREADYCALLED : BOOL;
	XLEAVESERVICESTATE : BOOL;
	XLEAVESERVICESTATEDISABLEDRIVE : BOOL;
	WLEAVESERVICESTATEPOWID : WORD;
	LRFOLLOWINGERRORACTIVE : LREAL;
	XMOTIONALLOWEDINACTUALSTATE : BOOL;
	XACTIVATEACTVALUESFORSYNCVALUES : BOOL;
	XCALLEDFROMINTERNALSTOP : BOOL;
	XCONNECTEDETCSLAVEDISABLED : BOOL;
	C_STRNOERROR : STRING := '-';
	C_STRUNDEFERROR : STRING := 'undefined';
	C_MAXFILTER : WORD := 2;
	C_MAXCOMP : WORD := 2;
	C_MAXFILTERINT : WORD := (c_MaxFilter + 1);
	C_UDILOGCOMPONENDID : UDINT := 16#2800;
	ACTACCELERATION : LREAL;
	ACTPOSITION : LREAL;
	ACTTORQUE : LREAL;
	ACTVELOCITY : LREAL;
	AXISID : DWORD;
	AXISPOOLCOUNT : WORD;
	AXISSLOT : L_MC1P_AxisSlot;
	AXISSTATE : L_MC1P_AXIS_STATE;
	CIA402ADVANCEDAXIS : BOOL;
	CMDCINH : BOOL;
	CMDFASTSTOP : BOOL;
	CMDFASTSTOPCINH : BOOL;
	CMDQSP : BOOL;
	CMDQSPCINH : BOOL;
	COMMANDEDPOSITION : LREAL;
	CYCLELENGTH : LREAL;
	DCTIMEACT : DWORD;
	DCTIMESET : DWORD;
	DCTIMESYNC : DWORD;
	DEVICE : L_MC1P_DriveType;
	DEVICECLASS : L_MC1P_DeviceClass;
	DRIVEENABLED : BOOL;
	DRIVEINITIALIZED : BOOL;
	DRVINFO : POINTER TO IIODrv.IoDrvInfo;
	ENCODERTYPE : L_Mc1P_EncoderType;
	FEEDCONSTANT : LREAL;
	GETACTIVELIMTERCONTROLWORD : DWORD;
	GETMASTERID : POINTER TO BYTE;
	HOMEPOSAVAILABLE : BOOL;
	HOMEPOSPERMANTENTSETACTIVE : BOOL;
	HOMEPOSPERMANTENTSETACTIVELOADENCODER : BOOL;
	ISVIRTUAL : BOOL;
	LICENSECONFIG : STRING;
	MODULEHANDLER : L_IMHP_IModuleHandler;
	NEWHOMEPOSLOADED : BOOL;
	QSPATFASTSTOPEND : BOOL;
	QSPWITHOUTREACTION : BOOL;
	RAMPDOWNINSERVICESTATE : BOOL;
	REAKTONMCFBERROR : BOOL;
	RESETFOLLOWINGERRORATFASTSTOPEND : BOOL;
	SELECTEDFORKINEMATIC : BOOL;
	SERVICEDIRECTION : L_MC1P_ServiceDirection;
	SETACCELERATIONFORSYNC : LREAL;
	SETHOMEPOSSTATEINDEPENDENTACTIVE : BOOL;
	SETPOSITIONFORSYNC : LREAL;
	SETPOSROUNDS : LREAL;
	SETTORQUEFORSYNC : LREAL;
	SETVELOCITYFORSYNC : LREAL;
	STARTPOSFORINTERNALSTOP : LREAL;
	STEADYSTATEID : DWORD;
	SUSPENDSWLIMITERRORREACTION : BOOL;
	TASKCYCLE : LREAL;
	TASKIDX : INT;
	TIMEDELAYACTPOS : LREAL;
	TIMEDELAYSETPOS : LREAL;
	TRANSMITCYCLESACTPOS : LREAL;
	TRAVERSINGRANGE : L_MC1P_TraversingRange;
	TRAVERSINGRANGEACT : L_MC1P_TraversingRange;
	USEDASINTERNALAXISINSTANCE : BOOL;
	USEDBYVIRTUALMASTER : BOOL;
END_VAR
END_FUNCTION_BLOCK

METHOD ACTIVATEACYCLICMODE
VAR_INPUT
	XACTIVATE : BOOL;
END_VAR
END_METHOD

METHOD CALCACTDIRECTION
END_METHOD

METHOD CALCACTPOSUNFILTERED : LREAL
END_METHOD

METHOD CALCSETDIRECTION : WORD
VAR_INPUT
	LRCYCVELIN : LREAL;
END_VAR
END_METHOD

METHOD CALLSIMULATION
VAR_INPUT
	CALLSTATE : L_UBUP_StateHandleCase;
END_VAR
END_METHOD

METHOD CHECKDIRECTION : BOOL
VAR_INPUT
	DIRECTION : MC_DIRECTION;
	ETYPEFUNCTION : L_MC1P_TypeFunction;
END_VAR
END_METHOD

METHOD CHECKMAXMODULOPOSDIFF
END_METHOD

METHOD CHECKPLNOTVALID : BOOL
END_METHOD

METHOD CHECKPLAUSIBILITYOFSETVALUES
END_METHOD

METHOD CHECKPOWER : BOOL
VAR_INPUT
	DWPOSSTATE : DWORD;
	LRVEL : LREAL;
END_VAR
END_METHOD

METHOD CHECKSLSVELOCITY : BOOL
END_METHOD

METHOD CHECKSETPOSINWINDOW : BOOL
END_METHOD

METHOD COMPENSATELOADPOSOFFSET
END_METHOD

METHOD ENABLEDRIVE : BOOL
VAR_INPUT
	XENABLE : BOOL;
END_VAR
END_METHOD

METHOD FLOATTOFRAC
VAR_INPUT
	LRINPUT : LREAL;
	PDIINTEGER : POINTER TO DINT;
	PUDIRESIDUAL : POINTER TO UDINT;
END_VAR
END_METHOD

METHOD FLOATTOFRACLINT
VAR_INPUT
	LRINPUT : LREAL;
	PLIINTEGER : POINTER TO LINT;
	PUDIRESIDUAL : POINTER TO UDINT;
END_VAR
END_METHOD

METHOD GENACTVALUES
END_METHOD

METHOD GETACTVEL : LREAL
END_METHOD

METHOD GETACTVELOCITYEXACT : LREAL
END_METHOD

METHOD GETACTIVEQUICKSTOPOPTION : L_MC1P_QuickStopOption
END_METHOD

METHOD GETAXISSLOT : UINT
END_METHOD

METHOD GETBRAKE : POINTER TO L_MC1P_BrakeControlBase
END_METHOD

METHOD GETBRAKESERVICE : POINTER TO L_MC1P_BrakeService
END_METHOD

METHOD GETCOUPLEDMASTERAXIS : POINTER TO BYTE
END_METHOD

METHOD GETCOUPLEDPHASINGMASTERAXIS : POINTER TO BYTE
END_METHOD

METHOD GETDRIVESTATE : BOOL
END_METHOD

METHOD GETEFFECTIVEMFESPEEDOFFSET : INT
VAR_INPUT
	INOFFSET : INT;
END_VAR
END_METHOD

METHOD GETMODULODIFF : LREAL
VAR_INPUT
	LRDIFF : LREAL;
END_VAR
VAR_IN_OUT
	AXIS : AXIS_REF;
END_VAR
END_METHOD

METHOD GETMODULOPOSITION : LREAL
VAR_INPUT
	LRNEWPOS : LREAL;
END_VAR
VAR_OUTPUT
	LRROUNDS : LREAL;
END_VAR
VAR_IN_OUT
	AXIS : AXIS_REF;
END_VAR
END_METHOD

METHOD GETPGMOVE : REFERENCE TO L_MC1P_PosProfiler
VAR_INPUT
	ITFPGACTIVE : L_MC1P_IPosProfilerActive;
END_VAR
END_METHOD

METHOD GETPGDUMMY : REFERENCE TO L_MC1P_PosProfiler
END_METHOD

METHOD GETPGSUPER : REFERENCE TO L_MC1P_PosProfiler
VAR_INPUT
	ITFPGACTIVE : L_MC1P_IPosProfilerActive;
END_VAR
END_METHOD

METHOD GETPHASESHIFT
VAR_OUTPUT
	LRPOS : LREAL;
	LRVEL : LREAL;
	LRACC : LREAL;
END_VAR
END_METHOD

METHOD GETPOINTERTOTPAXIS : POINTER TO _AXIS_REF_REAL
END_METHOD

METHOD GETRECEIVEDATA : DWORD
VAR_INPUT
	LWMASK : LWORD;
END_VAR
END_METHOD

METHOD GETTPWITHPOSITIONACTIVE : BOOL
VAR_INPUT
	SITPNUMBER : SINT;
END_VAR
END_METHOD

METHOD GETTPWITHTIMESTAMPACTIVE : BOOL
VAR_INPUT
	SITPNUMBER : SINT;
END_VAR
END_METHOD

METHOD HALTCALLEDBYABC
VAR_INPUT
	XCALLEDBYABC : BOOL;
END_VAR
END_METHOD

METHOD HLP_MODULOPOS : LREAL
VAR_INPUT
	LRPOSITION : LREAL;
	LRCYCLELENGTH : LREAL;
END_VAR
END_METHOD

METHOD HLP_MODULOPOS2 : LREAL
VAR_INPUT
	LRPOSITION : LREAL;
	LRCYCLELENGTH : LREAL;
	LRINVCYCLELENGTH : LREAL;
END_VAR
END_METHOD

METHOD INTOLERANCEWINDOW : BOOL
VAR_INPUT
	LRPOSITION : LREAL;
END_VAR
VAR_OUTPUT
	DIRECTION : MC_DIRECTION;
END_VAR
END_METHOD

METHOD INTERNALCONTROLMODE
END_METHOD

METHOD ISINCLUDEDINRECEIVEDATA : BOOL
VAR_INPUT
	LWMASK : LWORD;
END_VAR
END_METHOD

METHOD ISINCLUDEDINTRANSMITDATA : BOOL
VAR_INPUT
	LWMASK : LWORD;
END_VAR
END_METHOD

METHOD ISMOTIONALLOWED : BOOL
VAR_INPUT
	ETYPEFUNCTION : L_MC1P_TypeFunction;
END_VAR
VAR_IN_OUT
	XSUPERIMPOSED : BOOL;
END_VAR
END_METHOD

METHOD ISMOTIONALLOWED2 : BOOL
VAR_INPUT
	ETYPEFUNCTION : L_MC1P_TypeFunction;
	XCHECKHOMEPOS : BOOL;
END_VAR
VAR_OUTPUT
	EERRORCAUSE : L_IE1P_Error := L_IE1P_Error.NoError;
END_VAR
VAR_IN_OUT
	XSUPERIMPOSED : BOOL;
END_VAR
END_METHOD

METHOD LEAVESERVICESTATE
END_METHOD

METHOD LEAVESERVICESTATEBEAVIOUR : DINT
VAR_INPUT
	XDISABLEDRIVE : BOOL;
END_VAR
END_METHOD

METHOD LEAVESERVICESTATESTART : BOOL
END_METHOD

METHOD LIMITPROFILEDATA : WORD
VAR_INPUT
	PPROFLE : POINTER TO L_MC1P_ProfileParameter;
	PPROFLEOLD : POINTER TO L_MC1P_ProfileParameter;
END_VAR
END_METHOD

METHOD LOCKEDFORSINGLEMOTION
VAR_INPUT
	XLOCKED : BOOL;
END_VAR
END_METHOD

METHOD REGISTERAXESGROUP : BOOL
VAR_INPUT
	XUNREGISTER : BOOL;
	PAXESGROUP : POINTER TO BYTE;
END_VAR
END_METHOD

METHOD REGISTERFUNCTION : WORD
END_METHOD

METHOD REGISTERPHASINGFUNCTION : WORD
VAR_INPUT
	PMASTERAXIS : POINTER TO BYTE;
END_VAR
END_METHOD

METHOD REGISTERSUPERFUNCTION : WORD
END_METHOD

METHOD REGISTERSYNCFUNCTION : WORD
VAR_INPUT
	PMASTERAXIS : POINTER TO BYTE;
END_VAR
END_METHOD

METHOD RESETERRORSTATEOFCOMMANDS : BOOL
END_METHOD

METHOD RESETFOLLOWINGERROR
END_METHOD

METHOD RESETMOVEBUFFEREDINFO
END_METHOD

METHOD RESETMOVEINFO
END_METHOD

METHOD SERVICEMODEHANDLINGINDRIVEACTIVE : BOOL
END_METHOD

METHOD SETACTPOSITION
VAR_INPUT
	POSITION : LREAL;
	RELATIVE : BOOL;
END_VAR
END_METHOD

METHOD SETAXISSTATUSWORD
END_METHOD

METHOD SETBUFFERDATAALLOWED : BOOL
VAR_INPUT
	EMODE : MC_BUFFER_MODE;
	LRSPEED1 : LREAL;
	LRSPEED2 : LREAL;
	DWINSTANCE : __XWORD;
END_VAR
END_METHOD

METHOD SETDCBRAKE
VAR_INPUT
	XSETDCBRAKE : BOOL;
END_VAR
VAR_OUTPUT
	XDCBRAKEACTIVE : BOOL;
END_VAR
END_METHOD

METHOD SETENCODERITF
VAR_INPUT
	ENCODERIN : L_MC1P_IEncoderInterface;
END_VAR
END_METHOD

METHOD SETHOMEABSSWITCH
VAR_INPUT
	HOMEABSSWITCH : BOOL;
	XCHANGEDTOLOWLEVEL : BOOL;
END_VAR
END_METHOD

METHOD SETHOMEABSSWITCHOVERWRITE
VAR_INPUT
	XHOMEABSSWITCHSIGNAL : BOOL;
	XOVERWRITESIGNAL : BOOL;
END_VAR
END_METHOD

METHOD SETMACHINEDATA
END_METHOD

METHOD SETPHASESHIFT
VAR_INPUT
	LRPOS : LREAL;
	LRVEL : LREAL;
	LRACC : LREAL;
END_VAR
END_METHOD

METHOD SETPOSEQACTPOS
END_METHOD

METHOD SETPRECONTROLMODE
VAR_INPUT
	EPRECONTROLMODENEW : L_MC1P_PreControlMode := L_MC1P_PreControlMode.Automatic;
END_VAR
END_METHOD

METHOD SETTARGETPOS
VAR_INPUT
	LRTARGETPOSNEW : LREAL;
	LRTARGETPOSROUNDSNEW : LREAL;
	XVALID : BOOL;
END_VAR
END_METHOD

METHOD SETTARGETPOS2
VAR_INPUT
	LRTARGETPOSNEW : LREAL;
	LRTARGETPOSROUNDSNEW : LREAL;
	XVALID : BOOL;
	XRELMODE : BOOL;
END_VAR
END_METHOD

METHOD SETTORQUEVALUE
VAR_INPUT
	LRTORQUE : LREAL;
	WMODE : WORD;
END_VAR
END_METHOD

METHOD SETVELEQREFVALUE
VAR_INPUT
	LRREFVELOCITY : LREAL;
END_VAR
END_METHOD

METHOD SETVELOCITYOFFSET
VAR_INPUT
	WMODE : WORD;
	LROFFSETVELOCITY : LREAL;
END_VAR
END_METHOD

METHOD SPEEDEQZERO : BOOL
VAR_INPUT
	LRSPEEDIN : LREAL;
END_VAR
END_METHOD

METHOD SUSPENDFOLLOWINGERROR
VAR_INPUT
	XSUSPEND : BOOL;
END_VAR
END_METHOD

METHOD UPDATEERRORINFO
END_METHOD

METHOD UPDATEREADYFORMOTIONSTATUS : BOOL
VAR_INPUT
	AXISENABLED : BOOL;
END_VAR
END_METHOD

METHOD CALLRECIEVEPARAMETER
END_METHOD

METHOD CALLSDODATAHANDLING
END_METHOD

METHOD CALLTRANSMITPARAMETER
END_METHOD

METHOD CHECKCOMMUNCATION
END_METHOD

METHOD CHECKMAPPEDDATAVALID : BOOL
VAR_INPUT
	PADDDATA : POINTER TO BYTE;
	PDATA : POINTER TO POINTER TO BYTE;
END_VAR
VAR_OUTPUT
	XERROR : BOOL;
	EERRORID : L_IE1P_Error;
END_VAR
END_METHOD

METHOD GETMAPPEDDATA : POINTER TO BYTE
VAR_INPUT
	UIINDEX : WORD;
	USISUBINDEX : USINT;
	USISIZE : USINT;
	XWRITEACCESS : BOOL;
	PADDDATA : POINTER TO BYTE;
	PXWAITFORINITACCESS : POINTER TO BOOL;
END_VAR
VAR_OUTPUT
	EERRORID : L_IE1P_Error;
	XERROR : BOOL;
	USISIZEACT : USINT := 0;
END_VAR
END_METHOD

METHOD GETMAPPEDDATASUPPORT : BOOL
END_METHOD

METHOD RESETMAPPEDDATA
VAR_INPUT
	PADDDATA : POINTER TO BYTE;
END_VAR
END_METHOD

METHOD RESETSDODATA : DINT
VAR_INPUT
	IDX : DWORD;
	PDWSEMAPARACCESS : POINTER TO DWORD;
END_VAR
VAR_IN_OUT
	SDODATA : L_DCO_SdoData;
END_VAR
END_METHOD

METHOD CONFIGUREAXIS
END_METHOD

METHOD CONFIGUREAXIS2
END_METHOD

METHOD CONFIGUREAXISCONNECTOR
END_METHOD

METHOD CONFIGUREAXISCONNECTORBASICS : BOOL
END_METHOD

METHOD CONNECTCMDITFAUTOTUNING
END_METHOD

METHOD DETERMINETASKCYCLEINTERVAL : UDINT
END_METHOD

METHOD ENABLEAXISCONNECTOR : BOOL
END_METHOD

METHOD FINDANDCONNECTMOTIONUTILS
END_METHOD

METHOD GETTRANSMITCYCLESACTPOSFORPOSCTRL : LREAL
END_METHOD

METHOD REGISTERAXISPROPERTIES
END_METHOD

METHOD RESETAXISCONNECTOR
END_METHOD

METHOD SETAXISPROPERTIES
VAR_INPUT
	XUSEVIRTUAL : BOOL;
END_VAR
END_METHOD

METHOD UPDATEFATHERCONNECTOR
END_METHOD

METHOD CHECKAVAILABLECONTROLMODE : BOOL
END_METHOD

METHOD CONFIGURECONTROLMODE
VAR_OUTPUT
	EERRORID : L_IE1P_Error;
END_VAR
END_METHOD

METHOD GETDEFAULTCONTROLMODE : L_MC1P_ControlMode
END_METHOD

METHOD ISAVAILABLECONTROLMODE : BOOL
VAR_INPUT
	ECONTROLMODE : L_MC1P_ControlMode;
END_VAR
VAR_OUTPUT
	EERRORID : L_IE1P_Error;
END_VAR
END_METHOD

METHOD SETCONTROLMODE : BOOL
VAR_INPUT
	ECONTROLMODE : L_MC1P_ControlMode := L_MC1P_ControlMode.PosCtrlDrive;
	XKEEPACTPOSPRIORFDB : BOOL := FALSE;
	XRESTARTPOSITIONING : BOOL := FALSE;
END_VAR
VAR_OUTPUT
	EERRORID : L_IE1P_Error;
END_VAR
END_METHOD

METHOD SETCONTROLERITF
VAR_INPUT
	ITFCONTROLERNEW : L_MC1P_IControllerInterface;
END_VAR
END_METHOD

METHOD SETDEFAULTCONTROLMODE : BOOL
END_METHOD

METHOD CLEARERROR
VAR_INPUT
	PINSTANCE : POINTER TO BYTE := 0;
END_VAR
END_METHOD

METHOD CLEARERROR2
VAR_INPUT
	INSTANCEID : DWORD := 0;
END_VAR
END_METHOD

METHOD CLEARERRORID
VAR_INPUT
	PINSTANCE : POINTER TO BYTE := 0;
	WERRORID : WORD;
END_VAR
END_METHOD

METHOD CLEARERRORID2
VAR_INPUT
	INSTANCEID : DWORD := 0;
	WERRORID : WORD;
END_VAR
END_METHOD

METHOD CLEARERRORID3
VAR_INPUT
	INSTANCEID : DWORD := 0;
	WERRORID : WORD;
	DWEXTENDEDERRORINFO : DWORD;
END_VAR
END_METHOD

METHOD CLEARERRORINAXISSYSTEM
VAR_INPUT
	INSTANCEID : DWORD := 0;
END_VAR
END_METHOD

METHOD GETERRORITFID : DWORD
END_METHOD

METHOD HANDLEERRORENTRY : BOOL
VAR_INPUT
	WERRORID : L_IE1P_Error := 0;
	INSTANCEID : DWORD := 0;
	PSINSTANCENAME : POINTER TO BYTE := 0;
	DWEXTENDEDERRORINFO : DWORD;
	EERRORREACTION : L_IE1P_SeverityLevel := 0;
	XAUTORESET : BOOL;
	XNOLOGGINGENTRY : BOOL;
	XEXTERNALERROR : BOOL;
END_VAR
END_METHOD

METHOD NOTIFYERROR : BOOL
VAR_INPUT
	WERRORID : L_IE1P_Error := 0;
	PINSTANCE : POINTER TO BYTE := 0;
	PSINSTANCENAME : POINTER TO BYTE := 0;
	XSETERRORSTOP : BOOL := FALSE;
END_VAR
END_METHOD

METHOD NOTIFYERROR2 : BOOL
VAR_INPUT
	WERRORID : L_IE1P_Error := 0;
	INSTANCEID : DWORD := 0;
	PSINSTANCENAME : POINTER TO BYTE := 0;
	EERRORREACTION : L_IE1P_SeverityLevel := 0;
END_VAR
END_METHOD

METHOD NOTIFYERRORINAXISSYSTEM : BOOL
VAR_INPUT
	WERRORID : L_IE1P_Error := 0;
	INSTANCEID : DWORD := 0;
	PSINSTANCENAME : POINTER TO BYTE := 0;
	EERRORREACTION : L_IE1P_SeverityLevel := 0;
END_VAR
END_METHOD

METHOD SERERRORREACTIONEXTERN
VAR_INPUT
	EERRORREACTION : L_IE1P_SeverityLevel;
	WERRORID : WORD;
	INSTANCEID : DWORD := 0;
	XAUTORESET : BOOL;
	DWEXTENDEDERRORINFO : DWORD;
	XEXTERNALERROR : BOOL;
END_VAR
END_METHOD

METHOD UPDATEERRORREAKTION
VAR_INPUT
	SEVERITY : L_IE1P_SeverityLevel;
END_VAR
END_METHOD

METHOD EVENTCALLBACK : UDINT
VAR_INPUT
	PEVENTPARAM : POINTER TO EventParam;
END_VAR
END_METHOD

METHOD REGISTEREVENT
END_METHOD

METHOD UNREGISTEREVENT
END_METHOD

METHOD READMOTIONSTATE : BOOL
VAR_INPUT
	SOURCE : MC_SOURCE := MC_SOURCE.mcSetValue;
END_VAR
VAR_IN_OUT
	CONSTANTVELOCITY : BOOL;
	ACCELERATING : BOOL;
	DECELERATING : BOOL;
	DIRECTIONPOSITIVE : BOOL;
	DIRECTIONNEGATIVE : BOOL;
	INPOSITION : BOOL;
	STANDSTILLSETVELOCITY : BOOL;
	STANDSTILLACTVELOCITY : BOOL;
	ACTVELOCITYOLD : LREAL;
	SETVELOCITYOLD : LREAL;
	DRIVEENABLEDOLD : BOOL;
END_VAR
END_METHOD

METHOD ADDMASTERKINEMATIC : DINT
VAR_INPUT
	MASTER : L_MC1P_IKinematicMaster;
END_VAR
END_METHOD

METHOD ADDSLAVEKINEMATIC : DINT
VAR_INPUT
	SLAVE : L_MC1P_IKinematicSlave;
END_VAR
END_METHOD

METHOD COUPLEDAXISINERRORSTATE : BOOL
VAR_INPUT
	XCONTROLLEDSTOPPOSSIBLE : BOOL;
END_VAR
VAR_IN_OUT
	XSETQSP : BOOL;
	XSETCINH : BOOL;
END_VAR
END_METHOD

METHOD COUPLEDAXISSETERROR : BOOL
VAR_INPUT
	ESEVERITY : L_IE1P_SeverityLevel;
	WERRORID : WORD;
	DWEXTENDEDERRORINFO : DWORD;
END_VAR
END_METHOD

METHOD GANTRYSIGNALMONITORING : BOOL
END_METHOD

METHOD GETHOMINGDONESTATUS : BOOL
VAR_INPUT
	XDONE : BOOL;
END_VAR
END_METHOD

METHOD GETOPERATIONENABLEDSTATUS : BOOL
END_METHOD

METHOD HOMINGDONEOWNAXIS : BOOL
END_METHOD

METHOD HOMINGFINISH : BOOL
END_METHOD

METHOD HOMINGSETPARAMETER : BOOL
VAR_INPUT
	EHOMEMODE : L_MC1P_HomeMode;
	LRHOMEPOSITION : LREAL;
END_VAR
END_METHOD

METHOD HOMINGWAIT : BOOL
END_METHOD

METHOD ISMOTIONALLOWEDBYKIN : BOOL
VAR_INPUT
	ETYPEFUNCTION : L_MC1P_TypeFunction;
END_VAR
VAR_OUTPUT
	EERRORCAUSE : L_IE1P_Error := L_IE1P_Error.NoError;
END_VAR
END_METHOD

METHOD KINRESETPOSSIBLE : BOOL
END_METHOD

METHOD MOTIONALLOWEDINACTUALSTATE : BOOL
VAR_INPUT
	XALLOWED : BOOL;
END_VAR
END_METHOD

METHOD SETHOMINGDONE : DINT
VAR_INPUT
	XHOMINGDONE : BOOL;
END_VAR
END_METHOD

METHOD SLAVEABORTHOMING : DINT
END_METHOD

METHOD SLAVEDOHOMING : DINT
END_METHOD

METHOD SLAVEGENSETVALUES : DINT
END_METHOD

METHOD SLAVERESETERROR : BOOL
END_METHOD

METHOD SLAVERESETHOMEPOS : BOOL
VAR_INPUT
	ERESETINFO : L_IE1P_Error;
	XRESETPOSITION : BOOL;
END_VAR
END_METHOD

METHOD SLAVESETHOMEPOS : BOOL
VAR_INPUT
	POSITION : LREAL;
	RELATIVE : BOOL;
	XRESTARTPOSITIONING : BOOL := FALSE;
	EHOMEPOSINFO : L_IE1P_Error;
END_VAR
END_METHOD

METHOD GETINSTANCEANDTYPE : BOOL
VAR_OUTPUT
	PINSTANCEPOINTER : POINTER TO BYTE;
	EAXISTYPE : L_MC1P_AxisType;
END_VAR
END_METHOD

METHOD QUEUEDPARAMWRITINGACTIVE : BOOL
END_METHOD

METHOD RESETHOMEPOS
END_METHOD

METHOD RESETHOMEPOS2
VAR_INPUT
	ERESETINFO : L_IE1P_Error;
END_VAR
END_METHOD

METHOD RESETHOMEPOSLOADENCODER
VAR_INPUT
	ERESETINFO : L_IE1P_Error;
END_VAR
END_METHOD

METHOD SETHOMEPOSDEPENDONMODESTATEINDEPENDENT : BOOL
VAR_INPUT
	EHOMEMODE : L_MC1P_HomeMode;
	LRPOSITION : LREAL;
	LROFFSETPOSITION : LREAL;
	EHOMEPOSINFO : L_IE1P_Error;
END_VAR
VAR_OUTPUT
	XERROR : BOOL;
	EERRORID : L_IE1P_Error;
END_VAR
END_METHOD

METHOD SETHOMEPOSITION
VAR_INPUT
	POSITION : LREAL;
	RELATIVE : BOOL;
	XRESTARTPOSITIONING : BOOL := FALSE;
END_VAR
END_METHOD

METHOD SETHOMEPOSITION2
VAR_INPUT
	POSITION : LREAL;
	RELATIVE : BOOL;
	XRESTARTPOSITIONING : BOOL := FALSE;
	EHOMEPOSINFO : L_IE1P_Error;
END_VAR
END_METHOD

METHOD SETHOMEPOSITIONWITHMODROUNDS
VAR_INPUT
	POSITION : LREAL;
	RELATIVE : BOOL;
	ROUNDS : LREAL;
	XRESTARTPOSITIONING : BOOL;
	EHOMEPOSINFO : L_IE1P_Error;
END_VAR
END_METHOD

METHOD CALC_OUTPUTS
END_METHOD

METHOD CALC_STATUSSIGNALS
END_METHOD

METHOD ITFCHECKERRORRESETOCCURED : BOOL
VAR_IN_OUT
	RESETTIME : SYSTIME;
END_VAR
END_METHOD

METHOD ITFCLEARERROR : DWORD
VAR_INPUT
	ESEVERITY : L_IE1P_SeverityLevel;
	WERRORID : WORD;
	WCOMPID : WORD;
	DWINSTANCEID : DWORD := 0;
END_VAR
END_METHOD

METHOD ITFCLEARREACTION
VAR_INPUT
	EREACTION : L_IE1P_Reaction;
	DICLEARCOUNT : DINT;
	DWINSTANCEID : DWORD;
END_VAR
END_METHOD

METHOD ITFGETACTUALERRORCODE : DWORD
VAR_OUTPUT
	ESEVERITY : WORD;
END_VAR
END_METHOD

METHOD ITFREGISTERERRORINSTANCE : DWORD
END_METHOD

METHOD ITFRESETACTIVE : BOOL
END_METHOD

METHOD ITFRESETERROR : DWORD
VAR_INPUT
	ERRORHANDLE : SysTypes.RTS_IEC_HANDLE := 0;
END_VAR
END_METHOD

METHOD ITFRESETERRORREACTION
VAR_INPUT
	DWINSTANCEID : DWORD := 0;
END_VAR
END_METHOD

METHOD ITFSETERROR : DWORD
VAR_INPUT
	ESEVERITY : L_IE1P_SeverityLevel;
	WERRORID : WORD;
	WCOMPID : WORD;
	DWINSTANCEID : DWORD := 0;
	EREACTION : L_IE1P_Reaction;
END_VAR
END_METHOD

METHOD GETDIRECTION : WORD
VAR_INPUT
	VALUESOURCE : MC_SOURCE;
END_VAR
END_METHOD

METHOD GETMASTERERROR : BOOL
VAR_OUTPUT
	EERRORID : L_IE1P_Error;
END_VAR
END_METHOD

METHOD GETSTEADYSTATE : POINTER TO L_MC1P_SteadyState
END_METHOD

METHOD GETAXISFROMPOOL : POINTER TO AXIS_REF
VAR_INPUT
	WINDEX : WORD;
END_VAR
END_METHOD

METHOD CHECKINPOSITION
END_METHOD

METHOD SETINPOSITION
VAR_INPUT
	XDONE : BOOL;
	LRINTARGETPOSITION : LREAL;
END_VAR
END_METHOD

METHOD REQUESTINTERFACE : BOOL
VAR_INPUT
	ID : DINT;
	PITFUNKNOWN : POINTER TO L_UBUP_IUnknown;
END_VAR
END_METHOD

METHOD ACTIVATESS1
END_METHOD

METHOD CALCULATE_DECELERATION : LREAL
VAR_INPUT
	LRJERK : LREAL;
	LRTOTALTIME : LREAL;
	LRACTVEL : LREAL;
	LRTARGETVEL : LREAL;
	LRACCMAX : LREAL;
END_VAR
END_METHOD

METHOD CHECKLIMITERREQUESTS
END_METHOD

METHOD CHECKSLSCHANGES : BOOL
VAR_OUTPUT
	XLIMITERCONTROLCHANGED : BOOL;
	XSLSPARAMETERCHANGED : BOOL;
	XSLSNEWACTIVEDECELERATION : BOOL;
END_VAR
END_METHOD

METHOD CHECKSAFETYOPTIONAVAILABLE : BOOL
VAR_INPUT
	DWPRODUCTCODE : DWORD;
END_VAR
END_METHOD

METHOD LIMITSPEEDCONTROLLER
END_METHOD

METHOD PROCESSSSX
VAR_INPUT
	DWCONTROL : DWORD;
END_VAR
END_METHOD

METHOD UPDATEACTIVESLSSETVEL
VAR_INPUT
	LRVEL : LREAL;
END_VAR
END_METHOD

METHOD CHECKHWLIMITS : BOOL
END_METHOD

METHOD CHECKLIMITCHANGES : BOOL
VAR_OUTPUT
	XPOSSWLIMITCHANGED : BOOL;
	XNEGSWLIMITCHANGED : BOOL;
END_VAR
END_METHOD

METHOD CHECKMAXVALUES : BOOL
VAR_INPUT
	VELOCITY : LREAL;
	ACCELERATION : LREAL;
	JERK : LREAL;
END_VAR
END_METHOD

METHOD CHECKSWLIMITS : BOOL
VAR_INPUT
	XSETERRORSTOP : BOOL;
END_VAR
END_METHOD

METHOD DISABLESWLIMIT
VAR_INPUT
	XDISABLE : BOOL;
END_VAR
END_METHOD

METHOD GETACTDIRECTION : MC_DIRECTION
VAR_INPUT
	XCALCULATE : BOOL;
END_VAR
END_METHOD

METHOD GETSWLIMITSACTIVE : BOOL
END_METHOD

METHOD CALCCYCLELENGTH
END_METHOD

METHOD CALCULATESCALING : BOOL
END_METHOD

METHOD GETVIRTUAL : BOOL
END_METHOD

METHOD MACHINEDATACHANGED : BOOL
END_METHOD

METHOD WRITENEWMACHINEDATA
VAR_INPUT
	LRFEEDCONSTANTNEW : LREAL := 360.0;
	DWGEARDENOMINATORNEW : DWORD := 1;
	DWGEARNUMERATORNEW : DWORD := 1;
	DWADDGEARDENOMINATORNEW : DWORD := 1;
	DWADDGEARNUMERATORNEW : DWORD := 1;
	DWPOSRESOLUTIONNEW : DWORD := 65536;
	XORIENTATIONNEW : BOOL := FALSE;
	ETRAVERSINGRANGENEW : L_MC1P_TraversingRange := L_MC1P_TraversingRange.Limited;
	LRCYCLELENGTHNEW : LREAL := 360.0;
END_VAR
END_METHOD

METHOD COMPAREAXISNAME : BOOL
VAR_IN_OUT
	SAXISNAME : STRING;
END_VAR
END_METHOD

METHOD GETAXIS : POINTER TO AXIS_REF
END_METHOD

METHOD CALCSCALEFUNCTIONS
VAR_INPUT
	OFFSET : DWORD;
	INDEX : WORD;
END_VAR
END_METHOD

METHOD SETMACHINEDATAPARAMETER
END_METHOD

METHOD CALLCOMPFUNCTIONS
VAR_OUTPUT
	XCOMPERROR : BOOL;
END_VAR
END_METHOD

METHOD CALLFILTERFUNCTIONS
VAR_OUTPUT
	XFILTERERROR : BOOL;
END_VAR
END_METHOD

METHOD CHECKSETVALUESAVAILABLE
END_METHOD

METHOD RESETSETVALUESAVAILABLE
END_METHOD

METHOD RESTORESETVALUES
END_METHOD

METHOD SETCOMPITF : WORD
VAR_INPUT
	EINDEX : WORD;
	ITFCOMP : L_MC1P_ICompensationInterface;
END_VAR
END_METHOD

METHOD SETFILTERITF : WORD
VAR_INPUT
	EINDEX : WORD;
	ITFFILTER : L_MC1P_ISetvalueManipulationInterface;
	XFILTERINTERNALSET : BOOL;
END_VAR
END_METHOD

METHOD SETSETVALUESAVAILABLE
END_METHOD

METHOD SUSPENDSETVALUEFILTERCALL
VAR_INPUT
	XSUSPENDSETVALUEFILTERCALL : BOOL;
END_VAR
END_METHOD

METHOD ABORTACTIVEFUNCTION
END_METHOD

METHOD ACTIVATECOMPOFFSET : BOOL
VAR_INPUT
	EMODE : WORD := 0;
END_VAR
END_METHOD

METHOD COMPPOSOFFSET
VAR_INPUT
	EMODE : WORD := 0;
END_VAR
END_METHOD

METHOD COMPENSATETRANSMITCYCLES : BOOL
VAR_INPUT
	LRPOS : LREAL;
	LRVEL : LREAL;
	LRDELAYCYCLES : LREAL;
END_VAR
VAR_OUTPUT
	LRNEWPOS : LREAL;
	LRNEWVEL : LREAL;
	LRCORRECTION : LREAL;
END_VAR
END_METHOD

METHOD DRIVEQSP
END_METHOD

METHOD ERRORSTOP
END_METHOD

METHOD INTERNALSTOP : BOOL
VAR_INPUT
	XSTOP : BOOL;
	ESETSTATE : L_MC1P_AXIS_STATE;
	XPOSMODE : BOOL := FALSE;
	LRTARGETPOS : LREAL := 0;
	XABORTACTIVEFUNCTION : BOOL := TRUE;
END_VAR
VAR_IN_OUT
	XSTOPACTIVE : BOOL;
	XSTOPDONE : BOOL;
END_VAR
END_METHOD

METHOD MOVEBACKTOLASTSETPOS : BOOL
VAR_INPUT
	XSTOP : BOOL;
END_VAR
VAR_IN_OUT
	XSTOPACTIVE : BOOL;
	XSTOPDONE : BOOL;
END_VAR
END_METHOD

METHOD RAMPDOWN
END_METHOD

METHOD RAMPQSP
VAR_INPUT
	CALLEDFROMAPP : BOOL;
END_VAR
END_METHOD

METHOD RESETRAMPDOWN
END_METHOD

METHOD SETAXISSTOPINT : BOOL
VAR_INPUT
	XSTOP : BOOL;
	SCSTOPCMD : L_MC1P_StopOperation;
END_VAR
END_METHOD

METHOD SETFASTSTOPINT : BOOL
VAR_INPUT
	XSTOP : BOOL;
END_VAR
END_METHOD

METHOD SETSTANDSTILLSTATE
VAR_INPUT
	XRAMPDOWN : BOOL;
END_VAR
END_METHOD

METHOD STARTRAMPDOWN
END_METHOD

METHOD HLP_GETPARAMETER : BOOL
END_METHOD

METHOD HLP_GETPARAMETERPROPERTIES : BOOL
VAR_INPUT
	DIPARAMETER : DINT;
END_VAR
VAR_OUTPUT
	PPARAMADDR : POINTER TO BYTE := 0;
	EORDINALTYPE : L_MC1P_OrdinalType := L_MC1P_OrdinalType.otNONE;
	XREADWRITE : BOOL := FALSE;
	LRUNITFACTOR : LREAL := 1.0;
	LRDEFAULTVALUE : LREAL := 0.0;
	WVALUERANGES : WORD := 0;
	PVALUERANGES : POINTER TO L_MC1P_MinMaxValue := 0;
END_VAR
END_METHOD

METHOD HLP_INITPARREF
END_METHOD

METHOD HLP_READBOOLPARAMETER : BOOL
VAR_INPUT
	PARAMETER : DINT;
	PXVALUE : POINTER TO BOOL;
END_VAR
END_METHOD

METHOD HLP_READPARAMETER : BOOL
VAR_INPUT
	PARAMETER : DINT;
	PLRVALUE : POINTER TO LREAL;
END_VAR
END_METHOD

METHOD HLP_WRITEBOOLPARAMETER : BOOL
VAR_INPUT
	PARAMETER : DINT;
	PXVALUE : POINTER TO BOOL;
END_VAR
VAR_OUTPUT
	WERRORID : WORD;
END_VAR
END_METHOD

METHOD HLP_WRITEPARAMETER : BOOL
VAR_INPUT
	PARAMETER : DINT;
	PLRVALUE : POINTER TO LREAL;
END_VAR
VAR_OUTPUT
	WERRORID : WORD;
END_VAR
END_METHOD

METHOD AFTERREADINPUTS : INT
END_METHOD

METHOD AFTERWRITEOUTPUTS : INT
END_METHOD

METHOD BEFOREREADINPUTS : INT
END_METHOD

METHOD BEFOREWRITEOUTPUTS : INT
END_METHOD

METHOD CALCAFTERREADINPUTS : INT
END_METHOD

METHOD CALCAFTERWRITEOUTPUTS : INT
END_METHOD

METHOD CALCBEFOREREADINPUTS : INT
END_METHOD

METHOD CALCBEFOREWRITEOUTPUTS : INT
END_METHOD

METHOD FB_EXIT : BOOL
VAR_INPUT
	BINCOPYCODE : BOOL;
END_VAR
END_METHOD

METHOD INITFORSIMULATIONMODE : BOOL
VAR_INPUT
	WMODULETYPE : UINT;
	DWINSTANCE : UDINT;
	PCONNECTOR : POINTER TO IoConfigConnector;
END_VAR
END_METHOD

METHOD INITIALIZE : UDINT
VAR_INPUT
	WMODULETYPE : UINT;
	DWINSTANCE : UDINT;
	PCONNECTOR : POINTER TO IoConfigConnector;
END_VAR
END_METHOD

METHOD IODRVREADPARAMETER : UDINT
VAR_INPUT
	PCONNECTOR : POINTER TO IoConfigConnector;
	PPARAMETER : POINTER TO IoConfigParameter;
	PDATA : POINTER TO BYTE;
	DWBITSIZE : DWORD;
	DWBITOFFSET : DWORD;
END_VAR
END_METHOD

METHOD IODRVUPDATECONFIGURATION : UDINT
VAR_INPUT
	PCONNECTORLIST : POINTER TO IoConfigConnector;
	NCOUNT : DINT;
END_VAR
END_METHOD

METHOD IODRVUPDATEMAPPING : UDINT
VAR_INPUT
	PTASKMAPLIST : POINTER TO IoConfigTaskMap;
	NCOUNT : DINT;
END_VAR
END_METHOD

METHOD IODRVWRITEPARAMETER : UDINT
VAR_INPUT
	PCONNECTOR : POINTER TO IoConfigConnector;
	PPARAMETER : POINTER TO IoConfigParameter;
	PDATA : POINTER TO BYTE;
	DWBITSIZE : DWORD;
	DWBITOFFSET : DWORD;
END_VAR
END_METHOD

METHOD FB_INIT : BOOL
VAR_INPUT
	BINITRETAINS : BOOL;
	BINCOPYCODE : BOOL;
END_VAR
END_METHOD

METHOD FUNCTIONSUPPORTEDBYAXIS : BOOL
VAR_INPUT
	FUNID : L_MC1P_AxisFunction;
	XORIGINDEVICE : BOOL;
END_VAR
END_METHOD

METHOD GETDELAYFORFASTOUTPUTCALCULATION : LREAL
VAR_INPUT
	EVALUESOURCE : MC_SOURCE;
END_VAR
END_METHOD

METHOD GETINDEXOFENCODERCRC : WORD
END_METHOD

METHOD GETINDEXOFERRORCODE : DINT
END_METHOD

METHOD GETINDEXOFPOSCTRLADAPTVALUE
VAR_INPUT
	WSELECTION : WORD;
END_VAR
VAR_OUTPUT
	WINDEX : WORD;
	BYSUBINDEX : BYTE;
	BYSIZE : BYTE;
END_VAR
END_METHOD

METHOD GETINDEXOFSPEEDCTRLADAPTVALUE
VAR_INPUT
	WSELECTION : WORD;
END_VAR
VAR_OUTPUT
	WINDEX : WORD;
	BYSUBINDEX : BYTE;
	BYSIZE : BYTE;
END_VAR
END_METHOD

METHOD GETMAGNETISATIONFINISHED : BOOL
END_METHOD

METHOD GETMAXTORQUE : LREAL
END_METHOD

METHOD GETREFERENCETORQUE : LREAL
END_METHOD

METHOD GETTPDELAYFORFASTINPUTCALCULATION : LREAL
END_METHOD

METHOD GETVPPMAXVALUE : LREAL
END_METHOD

METHOD SETSPEEDCTRLLIMITATION : BOOL
VAR_INPUT
	XLIMIT : BOOL;
END_VAR
END_METHOD

METHOD SUPPORTLIMITSPEEDCONTROLLER : BOOL
VAR_OUTPUT
	WINDEX : WORD;
	BYSUBINDEX : BYTE;
	BYSIZE : BYTE;
END_VAR
END_METHOD

METHOD SUPPORTMFE : BOOL
END_METHOD

METHOD BRAKETESTDONEOWNAXIS : BOOL
END_METHOD

METHOD BRAKETESTFINISH : BOOL
END_METHOD

METHOD BRAKETESTWAIT : BOOL
END_METHOD

METHOD GETBTSTATUSFOLLOWER : LREAL
END_METHOD

METHOD GETBRAKETESTDONESTATUS : BOOL
VAR_INPUT
	XDONE : BOOL;
END_VAR
END_METHOD

METHOD SETBRAKETESTDONE : DINT
VAR_INPUT
	BRAKETESTDONE : BOOL;
END_VAR
END_METHOD

METHOD SLAVEABORTBRAKETEST : BOOL
VAR_INPUT
	XMAINABORTED : BOOL;
END_VAR
END_METHOD

METHOD SLAVEDOBRAKETEST : DINT
END_METHOD

METHOD GETGICYCLESFOLLOWER : LREAL
END_METHOD

METHOD GETGISTATUSFOLLOWER : LREAL
END_METHOD

METHOD GETGRINDINCYCLESDONE : WORD
VAR_INPUT
	WCYCLESIN : WORD;
END_VAR
END_METHOD

METHOD GETGRINDINDONESTATUS : BOOL
VAR_INPUT
	XDONE : BOOL;
END_VAR
END_METHOD

METHOD GRINDINDONEOWNAXIS : BOOL
END_METHOD

METHOD GRINDINFINISH : BOOL
END_METHOD

METHOD GRINDINPOW
VAR_INPUT
	XENABLE : BOOL;
	XDIRECTBRAKEMODE : BOOL := TRUE;
END_VAR
VAR_OUTPUT
	XEXTSTATUS : BOOL;
	XEXTVALID : BOOL;
END_VAR
END_METHOD

METHOD GRINDINWAIT : BOOL
END_METHOD

METHOD SETGIPOWID
VAR_INPUT
	WPOWID : WORD;
END_VAR
END_METHOD

METHOD SETGRINDINDONE : DINT
VAR_INPUT
	GRINDINDONE : BOOL;
END_VAR
END_METHOD

METHOD SLAVEABORTGRINDIN : BOOL
VAR_INPUT
	XMAINABORTED : BOOL;
END_VAR
END_METHOD

METHOD SLAVEDOGRINDIN : DINT
END_METHOD

METHOD CALCDISTANCE : LREAL
VAR_INPUT
	LRROUNDSACT : LREAL;
	LRROUNDSSET : LREAL;
	LRPOSACT : LREAL;
	LRPOSSET : LREAL;
END_VAR
VAR_IN_OUT
	AXIS : AXIS_REF;
END_VAR
END_METHOD

METHOD CALCTARGETPOS : LREAL
VAR_INPUT
	LRROUNDSACT : LREAL;
	LRROUNDSSET : LREAL;
	LRPOSACT : LREAL;
	LRPOSSET : LREAL;
END_VAR
VAR_OUTPUT
	EDIR : MC_DIRECTION;
END_VAR
VAR_IN_OUT
	AXIS : AXIS_REF;
END_VAR
END_METHOD

METHOD SETPOSRECOVERYDATA
VAR_INPUT
	XACTIVATE : BOOL;
	LRVEL : LREAL;
	LRACC : LREAL;
	LRDEC : LREAL;
	LRJERK : LREAL;
END_VAR
END_METHOD

(* ---- AXIS_REF_9400HL.pou ---- *)
FUNCTION_BLOCK AXIS_REF_9400HL EXTENDS _AXIS_REF_9400HL
VAR
	PARA_AXIS_REF_9400HL : L_MC1P_ParaInterface_AXIS_REF_9400HL;
END_VAR
END_FUNCTION_BLOCK

METHOD FB_INIT : BOOL
VAR_INPUT
	BINITRETAINS : BOOL;
	BINCOPYCODE : BOOL;
END_VAR
END_METHOD

(* ---- AXIS_REF_9400HL_CAN.pou ---- *)
FUNCTION_BLOCK AXIS_REF_9400HL_CAN EXTENDS _AXIS_REF_9400HL_CAN
VAR
	PARA_AXIS_REF_9400HL_CAN : L_MC1P_ParaInterface_AXIS_REF_9400HL_CAN;
END_VAR
END_FUNCTION_BLOCK

METHOD FB_INIT : BOOL
VAR_INPUT
	BINITRETAINS : BOOL;
	BINCOPYCODE : BOOL;
END_VAR
END_METHOD

(* ---- AXIS_REF_ENC_BPB.pou ---- *)
FUNCTION_BLOCK AXIS_REF_ENC_BPB EXTENDS _AXIS_REF_ENC_BPB
VAR
	PARA_AXIS_REF_ENC_BPB : L_MC1P_ParaInterface_AXIS_REF_ENC_BPB;
END_VAR
END_FUNCTION_BLOCK

METHOD FB_INIT : BOOL
VAR_INPUT
	BINITRETAINS : BOOL;
	BINCOPYCODE : BOOL;
END_VAR
END_METHOD

(* ---- AXIS_REF_ENC_FREE.pou ---- *)
FUNCTION_BLOCK AXIS_REF_ENC_FREE EXTENDS _AXIS_REF_ENC_FREE
VAR
	PARA_AXIS_REF_ENC_FREE : L_MC1P_ParaInterface_AXIS_REF_ENC_FREE;
END_VAR
END_FUNCTION_BLOCK

METHOD FB_INIT : BOOL
VAR_INPUT
	BINITRETAINS : BOOL;
	BINCOPYCODE : BOOL;
END_VAR
END_METHOD

(* ---- AXIS_REF_ENC_I500_ECAT.pou ---- *)
FUNCTION_BLOCK AXIS_REF_ENC_I500_ECAT EXTENDS _AXIS_REF_ENC_i500_ECAT
VAR
	PARA_AXIS_REF_ENC_I500_ECAT : L_MC1P_ParaInterface_AXIS_REF_ENC_i500_ECAT;
END_VAR
END_FUNCTION_BLOCK

METHOD FB_INIT : BOOL
VAR_INPUT
	BINITRETAINS : BOOL;
	BINCOPYCODE : BOOL;
END_VAR
END_METHOD

(* ---- AXIS_REF_ENC_I900_DRIVE.pou ---- *)
FUNCTION_BLOCK AXIS_REF_ENC_I900_DRIVE EXTENDS _AXIS_REF_ENC_i900_Target
VAR
	PARA_AXIS_REF_ENC_I900_DRIVE : L_MC1P_ParaInterface_AXIS_REF_ENC_i900_DRIVE;
END_VAR
END_FUNCTION_BLOCK

METHOD FB_INIT : BOOL
VAR_INPUT
	BINITRETAINS : BOOL;
	BINCOPYCODE : BOOL;
END_VAR
END_METHOD

(* ---- AXIS_REF_ENC_I900_DRIVE_CIA.pou ---- *)
FUNCTION_BLOCK AXIS_REF_ENC_I900_DRIVE_CIA EXTENDS _AXIS_REF_ENC_i900_CiA
VAR
	PARA_AXIS_REF_ENC_I900_DRIVE_CIA : L_MC1P_ParaInterface_AXIS_REF_ENC_i900_DRIVE_CIA;
END_VAR
END_FUNCTION_BLOCK

METHOD FB_INIT : BOOL
VAR_INPUT
	BINITRETAINS : BOOL;
	BINCOPYCODE : BOOL;
END_VAR
END_METHOD

(* ---- AXIS_REF_ENC_I900_ECAT.pou ---- *)
FUNCTION_BLOCK AXIS_REF_ENC_I900_ECAT EXTENDS _AXIS_REF_ENC_i900_ECAT
VAR
	PARA_AXIS_REF_ENC_I900_ECAT : L_MC1P_ParaInterface_AXIS_REF_ENC_i900_ECAT;
END_VAR
END_FUNCTION_BLOCK

METHOD FB_INIT : BOOL
VAR_INPUT
	BINITRETAINS : BOOL;
	BINCOPYCODE : BOOL;
END_VAR
END_METHOD

(* ---- AXIS_REF_ENC_IO_ETC.pou ---- *)
FUNCTION_BLOCK AXIS_REF_ENC_IO_ETC EXTENDS _AXIS_REF_ENC_IO_ETC
VAR
	PARA_AXIS_REF_ENC_IO_ETC : L_MC1P_ParaInterface_AXIS_REF_ENC_IO_ETC;
END_VAR
END_FUNCTION_BLOCK

METHOD FB_INIT : BOOL
VAR_INPUT
	BINITRETAINS : BOOL;
	BINCOPYCODE : BOOL;
END_VAR
END_METHOD

(* ---- AXIS_REF_ENC_UNIVERSAL.pou ---- *)
FUNCTION_BLOCK AXIS_REF_ENC_UNIVERSAL EXTENDS _AXIS_REF_Enc_Universal
VAR
	PARA_AXIS_REF_ENC_UNIVERSAL : L_MC1P_ParaInterface_AXIS_REF_ENC_UNIVERSAL;
END_VAR
END_FUNCTION_BLOCK

METHOD FB_INIT : BOOL
VAR_INPUT
	BINITRETAINS : BOOL;
	BINCOPYCODE : BOOL;
END_VAR
END_METHOD

(* ---- AXIS_REF_GENERIC.pou ---- *)
FUNCTION_BLOCK AXIS_REF_GENERIC EXTENDS _AXIS_REF_GENERIC
VAR
	PARA_AXIS_REF_GENERIC : L_MC1P_ParaInterface_AXIS_REF_GENERIC;
END_VAR
END_FUNCTION_BLOCK

METHOD FB_INIT : BOOL
VAR_INPUT
	BINITRETAINS : BOOL;
	BINCOPYCODE : BOOL;
END_VAR
END_METHOD

(* ---- AXIS_REF_I500_CAN.pou ---- *)
FUNCTION_BLOCK AXIS_REF_I500_CAN EXTENDS _AXIS_REF_i500_CAN
VAR
	PARA_AXIS_REF_I500_CAN : L_MC1P_ParaInterface_AXIS_REF_i500_CAN;
END_VAR
END_FUNCTION_BLOCK

METHOD FB_INIT : BOOL
VAR_INPUT
	BINITRETAINS : BOOL;
	BINCOPYCODE : BOOL;
END_VAR
END_METHOD

(* ---- AXIS_REF_I500_ETC.pou ---- *)
FUNCTION_BLOCK AXIS_REF_I500_ETC EXTENDS _AXIS_REF_i500_ETC
VAR
	PARA_AXIS_REF_I500_ETC : L_MC1P_ParaInterface_AXIS_REF_i500_ETC;
END_VAR
END_FUNCTION_BLOCK

METHOD FB_INIT : BOOL
VAR_INPUT
	BINITRETAINS : BOOL;
	BINCOPYCODE : BOOL;
END_VAR
END_METHOD

(* ---- AXIS_REF_I700.pou ---- *)
FUNCTION_BLOCK AXIS_REF_I700 EXTENDS _AXIS_REF_i700
VAR
	PARA_AXIS_REF_I700 : L_MC1P_ParaInterface_AXIS_REF_i700;
END_VAR
END_FUNCTION_BLOCK

METHOD FB_INIT : BOOL
VAR_INPUT
	BINITRETAINS : BOOL;
	BINCOPYCODE : BOOL;
END_VAR
END_METHOD
